(* IEC 61131-3 sources: daoli-st-library/DL_Algo (part 22) *)

(* ---- FB_DL_SortDiverterSeq.st ---- *)
(*
  DL Factory R83 | FB_DL_SortDiverterSeq
  功能：分拣分流器握手与故障恢复状态机，包裹到位后出分流指令并等动作确认、再等复位反馈，动作超时进重试（至多两次）后锁码，锁存可由复位沿解除恢复。
  开源溯源：无（clean-room 自研，依据公开工艺公式，来源=行业通用公式，许可证=MIT，借鉴点=公式结构）
  规则：R1-R21 全遵守
  ------------------------------------------------------------------
  分类 DL_Algo ｜ 复杂度 cx3 ｜ 版本 v1.0.0 ｜ 平台 纯 IEC 61131-3（TON、R_TRIG，无私有库）
  边界：一 本件只出分流指令与放行闸两路布尔命令，不驱动电磁阀线圈、不做包裹测速与到位判定（属主边界）；
        二 握手三段固定：到位（bParcelAt 上升沿）→ 分流指令（bDivertCmd）→ 动作确认（bAckFb 上升沿）
           → 复位反馈（bHomeFb 上升沿）→ 放行；三段证据齐全才置握手见证 _bHs；确认与复位反馈均为
           沿语义，须回零后再置位，电平自持不产生新沿（届时按超时走重试或锁码）；
        三 动作确认超时进重试：每次超时先把指令拉低（eRetry 相），重试间隔窗到再出指令；
           重试次数以 nMaxRetry 为预算（组态闸限定 0 至 2），预算耗尽仍超时即锁 402，不再重试；
        四 复位反馈超时锁 403；到位滞留超时锁 404；组态或预算越域锁 401；非法相位锁 405；
           故障锁存由 bReset 上升沿解除（唯一解除路径，R188），锁存期码位一律回放（R152）；
        五 R510 守卫（默认引脚值组合不得绕过握手直达放行）：放行闸为 _bHandshakeSeen 与相位、下游许可、
           使能与锁存位的合取式，默认引脚组合（bParcelAt、bAckFb、bHomeFb、bDownstreamClear 全假）下
           握手见证位恒假，放行闸结构上恒闭；另设「eDone 相缺握手见证即判非法相位」的防御性拦截行；
           本场景不加新码（R90 反证：默认组合下无任何输出组合能把放行闸观测为真，故无需独立码位稀释预留带）；
        六 每相一个专属定时器（到位滞留、动作确认、复位反馈、重试间隔），IN 只串本相使能与锁存闸，
           相迁移即 IN 归假并自复位（R18）；四窗分属不同相、无同拍双窗，R100 配比约束不适用；
        七 单向计数纪律（R45 ③）：重试计数 _nRetry 的自增点唯一（eCmd 超时分支），其余位置只做清零；
           零点共有三处且互斥（首扫与复位沿、eIdle 迁出、eDone 迁出），无任何递减路径；
        八 无全局变量、无外部变量声明、无物理地址寻址。
  输出契约：bDivertCmd 为分流指令电平（仅 eCmd 相，故障与失能一律归零）；bReleaseGate 为放行闸；
        bHandshakeOk 为握手见证位（三段证据齐全，新循环起点清零）；nRetryCnt 为已用重试次数；
        bDone 为保持式完成位（包裹离开时清零，R28 5.9 清零点）；iErrCode 为锁存回放。
  修订记录：2026-11-24 v1.0.0 R83 首版（批 R83 · 序号 40）
*)

TYPE E_DL_SdvPhase :
(
    eIdle  := 0,  // 空闲等使能 / idle, waiting for the enable
    eWait  := 10, // 等到位：等包裹到位沿 / waiting for the parcel arrival edge
    eCmd   := 20, // 分流指令：出指令并等动作确认 / the divert command is on and the acknowledgement is awaited
    eBack  := 30, // 等复位：等分流器复位反馈 / waiting for the diverter home feedback
    eRetry := 40, // 重试：指令拉低，等重试间隔窗 / retrying, the command is off while the gap window runs
    eDone  := 50, // 完成：握手齐全，等包裹离开后放行结束 / done, the handshake is complete and the parcel leaves
    eFault := 90  // 故障：成因锁存等复位沿 / fault, the cause is latched until the reset edge
);
END_TYPE

TYPE E_DL_SdvCause :
(
    eNone     := 0, // 无成因 / no cause
    eCfgBad   := 1, // 组态或重试预算越域（故障级，与 bError 配对）/ the configuration or the retry budget is out of domain, fault grade paired with bError
    eAckTo    := 2, // 动作确认超时且预算耗尽（故障级，与 bError 配对）/ the acknowledgement timed out with the budget exhausted, fault grade paired with bError
    eHomeTo   := 3, // 复位反馈超时（故障级，与 bError 配对）/ the home feedback timed out, fault grade paired with bError
    eWaitTo   := 4, // 包裹到位滞留超时（故障级，与 bError 配对）/ the parcel arrival lingered past its window, fault grade paired with bError
    ePhaseBad := 5  // 非法相位或缺握手见证的完成相（故障级，与 bError 配对）/ an illegal phase or a done phase without the handshake witness, fault grade paired with bError
);
END_TYPE

FUNCTION_BLOCK FB_DL_SortDiverterSeq
VAR CONSTANT
    DL_SDV_RETRY_MAX : INT := 2; // 重试次数硬上限（预算域上限）[次] / the hard upper bound of the retry budget [time]
END_VAR
VAR_INPUT
    bEnable          : BOOL := TRUE;  // 使能，失能回空闲且指令归零 [-] / enable, a disable returns to idle with the command zeroed
    bReset           : BOOL := FALSE; // 复位上升沿清故障锁存并回空闲 [-] / reset rising edge clears the latch and returns to idle
    bParcelAt        : BOOL := FALSE; // 包裹到位光电（上升沿起握手）[-]/ the parcel arrival photo sensor, its rising edge starts the handshake
    bAckFb           : BOOL := FALSE; // 分流器动作确认反馈（上升沿）[-]/ the diverter action acknowledgement, its rising edge
    bHomeFb          : BOOL := FALSE; // 分流器复位反馈（上升沿）[-]/ the diverter home feedback, its rising edge
    bDownstreamClear : BOOL := FALSE; // 下游放行许可（默认假，保守侧）[-]/ the downstream clearance, default false on the safe side
    nMaxRetry        : INT := 2;      // 允许重试次数（域 0 至 2）[次] / the allowed retry count, domain zero to two [time]
    tWaitTo          : TIME := T#10S; // 包裹到位滞留超时窗 [毫秒] / the parcel arrival lingering window [millisecond]
    tAckTo           : TIME := T#2S;  // 动作确认超时窗 [毫秒] / the acknowledgement timeout window [millisecond]
    tHomeTo          : TIME := T#5S;  // 复位反馈超时窗 [毫秒] / the home feedback timeout window [millisecond]
    tRetryGap        : TIME := T#1S;  // 重试间隔窗（指令拉低时段）[毫秒] / the retry gap window while the command is off [millisecond]
END_VAR
VAR_OUTPUT
    bBusy        : BOOL := FALSE; // 本包裹处理中 [-] / a parcel is being handled
    bDone        : BOOL := FALSE; // 本包裹握手齐全（保持式，包裹离开清零）[-] / the handshake completed for this parcel
    bFault       : BOOL := FALSE; // 故障锁存 [-] / the fault latch
    bError       : BOOL := FALSE; // 故障标志，与锁存位同源 [-] / the fault flag sharing the latch source
    iErrCode     : INT := 0;      // 错误码（锁存回放，复位沿清零）[码] / the error code replayed from the latch [code]
    ePhase       : E_DL_SdvPhase := E_DL_SdvPhase.eIdle; // 相位出口 [枚举] / the phase outlet [enum]
    bDivertCmd   : BOOL := FALSE; // 分流指令电平（仅 eCmd 相）[-] / the divert command level, eCmd only
    bReleaseGate : BOOL := FALSE; // 放行闸（握手齐全且下游许可）[-] / the release gate, handshake complete and downstream clear
    bHandshakeOk : BOOL := FALSE; // 握手见证位（三段证据齐全）[-] / the handshake witness covering all three evidences
    nRetryCnt    : INT := 0;      // 已用重试次数 [次] / the used retry count [time]
END_VAR
VAR
    rtReset    : R_TRIG; // 复位沿，段 2 无条件刷新 / the reset edge, refreshed unconditionally
    rtParcel   : R_TRIG; // 包裹到位沿，段 2 无条件刷新 / the parcel arrival edge, refreshed unconditionally
    rtAck      : R_TRIG; // 动作确认沿，段 2 无条件刷新 / the acknowledgement edge, refreshed unconditionally
    rtHome     : R_TRIG; // 复位反馈沿，段 2 无条件刷新 / the home feedback edge, refreshed unconditionally
    tonWait    : TON;    // 到位滞留超时窗，只串 eWait 相 / the arrival lingering window gated by eWait
    tonAck     : TON;    // 动作确认超时窗，只串 eCmd 相 / the acknowledgement timeout gated by eCmd
    tonHome    : TON;    // 复位反馈超时窗，只串 eBack 相 / the home feedback timeout gated by eBack
    tonRetry   : TON;    // 重试间隔窗，只串 eRetry 相 / the retry gap window gated by eRetry
    _ePhase    : E_DL_SdvPhase := E_DL_SdvPhase.eIdle; // 内部相位，CASE 唯一写入目标 / the internal phase, the only CASE target
    _eCause    : E_DL_SdvCause := E_DL_SdvCause.eNone; // 故障级成因，锁存至复位沿 / the fault cause latched until reset
    _bFault    : BOOL := FALSE; // 故障锁存位 [-] / the fault latch
    _iErrLch   : INT := 0;      // 码位锁存槽（复位沿清零）[码] / the latched code, cleared at the reset edge
    _bDone     : BOOL := FALSE; // 完成位内部锁存（清零归属：段 3 复位沿与 eDone 迁出分支）[-] / the internal done bit
    _bHs       : BOOL := FALSE; // 握手见证位内部锁存（三段证据齐全，新循环起点清零）[-] / the handshake witness, cleared at a new cycle
    _bInit     : BOOL := FALSE; // 首扫初始化完成标志（R310）[-] / the first scan initialisation flag
    _bCfgOk    : BOOL := FALSE; // 组态与重试预算域内 [-] / the configuration and the retry budget are inside their domain
    _nRetry    : INT := 0;      // 已用重试次数（单点自增，R45 ③）[次] / the used retry count, incremented at one point only [time]
END_VAR
// 段 0｜组态与重试预算域闸：参与判据换算的引脚逐项枚举（R151）
_bCfgOk := (nMaxRetry >= 0) AND (nMaxRetry <= DL_SDV_RETRY_MAX) // 重试预算落在 [0, 硬上限] / the retry budget inside its domain
    AND (tWaitTo > T#0S) AND (tAckTo > T#0S) AND (tHomeTo > T#0S) AND (tRetryGap > T#0S); // 四个时间引脚域闸 / the four time pins domain gate
// 段 1｜定时器与沿检测无条件周期刷新，IN 只串本相使能与锁存闸（R7、R18）
rtReset(CLK := bReset); // 复位沿无条件刷新 / unconditional refresh of the reset edge
rtParcel(CLK := bParcelAt); // 包裹到位沿无条件刷新 / unconditional refresh of the parcel arrival edge
rtAck(CLK := bAckFb); // 动作确认沿无条件刷新 / unconditional refresh of the acknowledgement edge
rtHome(CLK := bHomeFb); // 复位反馈沿无条件刷新 / unconditional refresh of the home feedback edge
tonWait(IN := (_ePhase = E_DL_SdvPhase.eWait) AND bParcelAt AND (NOT _bFault), PT := tWaitTo); // 到位滞留窗：只串 eWait 相且到位光电为电平（空载等待不计时）/ the arrival window gated by eWait and the live photo level
tonAck(IN := (_ePhase = E_DL_SdvPhase.eCmd) AND (NOT _bFault), PT := tAckTo); // 动作确认窗，只串 eCmd 相 / the acknowledgement window gated by eCmd only
tonHome(IN := (_ePhase = E_DL_SdvPhase.eBack) AND (NOT _bFault), PT := tHomeTo); // 复位反馈窗，只串 eBack 相 / the home window gated by eBack only
tonRetry(IN := (_ePhase = E_DL_SdvPhase.eRetry) AND (NOT _bFault), PT := tRetryGap); // 重试间隔窗，只串 eRetry 相 / the retry gap gated by eRetry only
// 段 2｜首扫初始化与复位沿同块，作用域逐项声明（R310、R311）
IF (NOT _bInit) OR rtReset.Q THEN // 首扫一拍或复位沿 / the first scan or the reset edge
    _bInit := TRUE; // 首扫完成标志（复位沿重复置位同效）/ the first scan flag, the same effect on reset
    _bFault := FALSE; _eCause := E_DL_SdvCause.eNone; _iErrLch := 0; // 作用域一：清锁存、清成因、清码位槽 / scope one, clear the latch, the cause and the code
    _bDone := FALSE; _bHs := FALSE; _ePhase := E_DL_SdvPhase.eIdle; // 作用域二：清完成位、清握手见证并迁回空闲 / scope two, clear done and the witness and migrate to idle
    _nRetry := 0; // 作用域三：清重试计数（三处清零点之一，另两处为 eIdle 与 eDone 迁出）/ scope three, clear the retry counter, one of three clear points
END_IF
// 段 3｜故障判据与锁存：未锁存才判，锁存与迁相同拍执行（R107、FB50-1④、R152）
IF NOT _bFault THEN // 未锁存才判，锁存后一律回放 / judge only while unlatched
    IF NOT _bCfgOk THEN // 组态或重试预算越域 / the configuration or the retry budget is out of domain
        _eCause := E_DL_SdvCause.eCfgBad; _iErrLch := 401; bError := TRUE; // 故障级成因、码位与标志（R45 配对）
        _bFault := TRUE; _ePhase := E_DL_SdvPhase.eFault; // 置锁存并同拍迁故障相 / latch and migrate in the same scan
    ELSIF (_ePhase = E_DL_SdvPhase.eDone) AND (NOT _bHs) THEN // R510 守卫：完成相缺握手见证即判非法（防御性拦截，结构上不可达）
        _eCause := E_DL_SdvCause.ePhaseBad; _iErrLch := 405; bError := TRUE; // 故障级成因、码位与标志（R45 配对）
        _bFault := TRUE; _ePhase := E_DL_SdvPhase.eFault; // 置锁存并同拍迁故障相 / latch and migrate in the same scan
    END_IF
END_IF
// 段 4｜相位状态机：ENUM ＋ CASE ＋ ELSE 非法相位兜底（R6、R128）
CASE _ePhase OF
E_DL_SdvPhase.eIdle: // 空闲相：退出条件二（使能给出、使能未给则驻留）
    IF bEnable THEN // 使能给出 / the enable is given
        _nRetry := 0; _bHs := FALSE; _ePhase := E_DL_SdvPhase.eWait; // 清重试与见证并迁等到位相 / clear the retry and the witness and migrate to wait
    END_IF
E_DL_SdvPhase.eWait: // 等到位相：退出条件三（到位沿、滞留超时、使能丢失）
    IF NOT bEnable THEN // 使能丢失 / the enable was lost
        _ePhase := E_DL_SdvPhase.eIdle; // 回空闲 / back to idle
    ELSIF rtParcel.Q THEN // 到位沿先消化（拍 N 进入：本相起点、本拍行为：拒绝出指令、拍 N+1 转出：指令相）
        _ePhase := E_DL_SdvPhase.eCmd; // 迁分流指令相 / migrate to the command phase
    ELSIF tonWait.Q THEN // 到位光电长期为真而无上升沿（包裹卡滞）/ the photo stayed true without an edge, the parcel is stuck
        _eCause := E_DL_SdvCause.eWaitTo; _iErrLch := 404; bError := TRUE; // 故障级成因、码位与标志（R45 配对）
        _bFault := TRUE; _ePhase := E_DL_SdvPhase.eFault; // 置锁存并迁故障相 / latch and migrate to the fault phase
    END_IF
E_DL_SdvPhase.eCmd: // 分流指令相：指令保持，退出条件三（确认沿、确认超时、使能丢失），事件优先于超时（R275）
    IF NOT bEnable THEN // 使能丢失 / the enable was lost
        _ePhase := E_DL_SdvPhase.eIdle; // 回空闲（指令归零由出口执行）/ back to idle, the outlet zeroes the command
    ELSIF rtAck.Q THEN // 动作确认沿先消化 / digest the acknowledgement edge first
        _ePhase := E_DL_SdvPhase.eBack; // 迁等复位相 / migrate to the home phase
    ELSIF tonAck.Q THEN // 动作确认超时 / the acknowledgement timed out
        IF _nRetry < nMaxRetry THEN // 预算内：进重试 / inside the budget, retry
            _nRetry := _nRetry + 1; // 重试计数单点自增（R45 ③）/ the single increment point of the retry counter
            _ePhase := E_DL_SdvPhase.eRetry; // 迁重试相（指令拉低等间隔窗）/ migrate to retry with the command off
        ELSE // 预算耗尽：锁码 / the budget is exhausted, latch the code
            _eCause := E_DL_SdvCause.eAckTo; _iErrLch := 402; bError := TRUE; // 故障级成因、码位与标志（R45 配对）
            _bFault := TRUE; _ePhase := E_DL_SdvPhase.eFault; // 置锁存并迁故障相 / latch and migrate to the fault phase
        END_IF
    END_IF
E_DL_SdvPhase.eBack: // 等复位相：退出条件三（复位沿、复位超时、使能丢失）；复位沿即三段证据齐全
    IF NOT bEnable THEN // 使能丢失 / the enable was lost
        _ePhase := E_DL_SdvPhase.eIdle; // 回空闲 / back to idle
    ELSIF rtHome.Q THEN // 复位反馈沿：置握手见证并转完成 / the home edge completes the handshake
        _bHs := TRUE; _bDone := TRUE; _ePhase := E_DL_SdvPhase.eDone; // 置见证位与完成位并迁完成相 / raise the witness and done and migrate
    ELSIF tonHome.Q THEN // 复位反馈超时 / the home feedback timed out
        _eCause := E_DL_SdvCause.eHomeTo; _iErrLch := 403; bError := TRUE; // 故障级成因、码位与标志（R45 配对）
        _bFault := TRUE; _ePhase := E_DL_SdvPhase.eFault; // 置锁存并迁故障相 / latch and migrate to the fault phase
    END_IF
E_DL_SdvPhase.eRetry: // 重试相：指令拉低，退出条件二（间隔窗到期回指令相、使能丢失回空闲）
    IF NOT bEnable THEN // 使能丢失 / the enable was lost
        _ePhase := E_DL_SdvPhase.eIdle; // 回空闲 / back to idle
    ELSIF tonRetry.Q THEN // 重试间隔窗到期 / the retry gap expired
        _ePhase := E_DL_SdvPhase.eCmd; // 回指令相重新出指令 / back to the command phase
    END_IF
E_DL_SdvPhase.eDone: // 完成相：退出条件二（包裹离开、使能丢失），完成位与见证位在此清零（单一清零点）
    IF (NOT bParcelAt) OR (NOT bEnable) THEN // 包裹离开或失能 / the parcel left or the enable was lost
        _bDone := FALSE; _bHs := FALSE; _nRetry := 0; _ePhase := E_DL_SdvPhase.eIdle; // 清完成位、见证位与重试并回空闲 / clear done, the witness and the retry and return to idle
    END_IF
E_DL_SdvPhase.eFault: // 故障相：成因锁存回放，唯一解除路径为 bReset 上升沿（R188）
    IF NOT bEnable THEN _ePhase := E_DL_SdvPhase.eIdle; END_IF // 失能迁空闲（锁存位仍须复位沿解除）/ migrate to idle, the latch still needs the reset edge
ELSE // 非法相位兜底（R6、R128）/ the illegal phase fallback
    _eCause := E_DL_SdvCause.ePhaseBad; _iErrLch := 405; bError := TRUE; // 故障级成因、码位与标志（R45 配对）
    _bFault := TRUE; _ePhase := E_DL_SdvPhase.eFault; // 置锁存并迁故障相 / latch and migrate to the fault phase
END_CASE
IF _bFault AND (_ePhase <> E_DL_SdvPhase.eFault) THEN // 段尾迁移闸：任何锁存路径不得留在业务相（FB50-1④）
    _ePhase := E_DL_SdvPhase.eFault; // 统一迁故障相 / force the fault phase
END_IF
// 段 5｜统一出口：指令与放行闸单点映射，R510 守卫在放行闸结构上落地
bDivertCmd := (_ePhase = E_DL_SdvPhase.eCmd) AND bEnable AND (NOT _bFault); // 分流指令：仅指令相且未失能未锁存 / the divert command only in the command phase while enabled and unlatched
bReleaseGate := _bHs AND (_ePhase = E_DL_SdvPhase.eDone) AND bDownstreamClear AND bEnable AND (NOT _bFault); // 放行闸：握手见证与相位、下游许可、使能、锁存位五者合取（默认组合下恒闭，R510 守卫）
bHandshakeOk := _bHs; // 握手见证位单点映射 / single point mapping of the handshake witness
nRetryCnt := _nRetry; // 重试计数单点映射 / single point mapping of the retry counter
bBusy := bEnable AND (_ePhase <> E_DL_SdvPhase.eIdle) AND (_ePhase <> E_DL_SdvPhase.eDone) AND (_ePhase <> E_DL_SdvPhase.eFault); // 运行位排除空闲完成与故障 / the busy bit excludes idle, done and fault
bDone := _bDone; // 完成位单点映射（保持式）/ single point mapping of the held done bit
bFault := _bFault; // 故障锁存单点映射 / single point mapping of the latch
IF _bFault THEN // 故障期回放锁存码，不在故障相按当下输入重推（R152）/ replay the latched code
    iErrCode := _iErrLch; bError := TRUE; // 锁存码回放、故障标志同源 / replay the code and share the latch source
ELSE // 非故障期 / outside fault
    iErrCode := 0; bError := FALSE; // 无故障码与无故障标志 / no code and no flag
END_IF
ePhase := _ePhase; // 相位出口单点映射 / single point mapping of the phase
END_FUNCTION_BLOCK

(* ---- FB_DL_SplitRangeControl.st ---- *)
(*==============================================================================
 * 组件名称 (Component)  : FB_DL_SplitRangeControl
 * 所属子库 (Sublibrary) : DL_Algo
 * 当前版本 (Version)    : 1.0.0
 * 兼容性   (Platform)   : CODESYS 3.5 / TwinCAT 3 / 汇川 InoProShop / Machine Expert
 *                         仅依赖纯 IEC 61131-3 数学运算，零库依赖，零厂商方言
 * 功能描述 (Function)   : 分程输出分配。把单一控制器输出（-100..100%）分配为
 *                         两路执行器信号：正半区驱动加热通道、负半区驱动冷却
 *                         通道，中央死区间隙防双阀同开；两路输出各自按独立量程
 *                         二次映射，支持加热通道反相。现场用途：温控冷热双执
 *                         行器、蒸汽 / 冷水阀对。
 * 开源溯源 (Origin)     : 原创实现。分程控制功能分类与参数域参考过程控制经典
 *                         文献（split-range pairing）的公开语义描述，
 *                         未复制任何厂商源码，clean-room 重写。
 * 本文件内含       : TYPE  E_DL_SplitState（配套枚举，归属 DL_Algo）
 *                    FB    FB_DL_SplitRangeControl
 * 依赖     (Depends)    : 无 DL_ 内部依赖；Standard.library 无实例依赖
 * 红线自检 (Redline)    : R1 ✓ 零全局变量表与外部变量引用 ｜ R2 ✓ 零物理 IO 地址直写
 *                         R3 ✓ 纯 IEC 61131-3 ｜ R4 ✓ 防除零+钳位+非有限值防御
 *                         R5 ✓ 全变量中英双语同行注释 ｜ R6 ✓ 五态 ENUM+CASE+ELSE
 *                         R7 ✓ 本块无定时器 / 边沿实例（无可刷新项，天然合规）
 * 修订历史 (Revision)   :
 *   2026-11-15  v1.0.0  首版入库 · Round 04 · Level 1 DL_Algo
 * 验收向量 (Acceptance) :
 *   V1 正半区：fCtrlIn=50 → fOutHeat=50、fOutCool=0、bHeatActive=TRUE
 *   V2 负半区：fCtrlIn=-40 → fOutCool=40、fOutHeat=0、bCoolActive=TRUE
 *   V3 死区：fCtrlIn=1.0 且 fGap=2.0 → 两路输出均为 0
 *   V4 反相：fCtrlIn=50 且 bInvertHeat=TRUE → fOutHeat=50 映射后取 100-x
 *   V5 非有限值：fCtrlIn 写入非法浮点 → 两路输出保持上一拍且码 0002_0004
 *   V6 二次映射：rOutHeatMin=20 → fOutHeat 从 20 起算
 *============================================================================*)

(*-----------------------------------------------------------------------------
 * 枚举: E_DL_SplitState（归属 DL_Algo，与 FB_DL_SplitRangeControl 同文件）
 * 含义: 分程分配离散状态。数值步长留空位便于后续插态而不破坏已有工程。
 *----------------------------------------------------------------------------*)
TYPE E_DL_SplitState :
(
    eIdle     := 0,    // 使能关：两路输出回各自量程下限 / Idle: enable off, both outputs at range low
    eHeatZone := 10,   // 加热区：正半区驱动加热通道 / Heat zone: positive half drives heating channel
    eDeadband := 20,   // 中央死区：两路输出均为零 / Central deadband: both outputs zero
    eCoolZone := 30,   // 冷却区：负半区驱动冷却通道 / Cool zone: negative half drives cooling channel
    eFault    := 99    // 故障兜底态：非法状态进入，输出安全值 / Fault fallback: illegal state, safe output
);
END_TYPE

(*==============================================================================
 * 功能块: FB_DL_SplitRangeControl
 * 调用约定: 每个扫描周期无条件调用一次。
 * 无状态泄漏: 全部状态驻留于实例私有 VAR，零全局引用，可多实例并行。
 * 工程披露: tSampleTime 仅用于与子库其余组件保持引脚一致性与未来扩展。
 *============================================================================*)
FUNCTION_BLOCK FB_DL_SplitRangeControl
VAR_INPUT
    bEnable     : BOOL := FALSE;      // 总使能，FALSE 时两路回量程下限 / Master enable, FALSE drives both to range low
    fCtrlIn     : REAL := 0.0;        // 控制器输入 [%]，-100..100 / Controller input in percent, -100..100
    fGap        : REAL := 2.0;        // 中央死区 [%]，负值钳 0 / Central deadband in percent, negative clamped
    rCtrlMax    : REAL := 100.0;      // 输入满量程幅值 [%]，须大于 0 / Input full-scale magnitude in percent
    rOutHeatMin : REAL := 0.0;        // 加热通道输出下限 [%] / Heating channel output lower limit
    rOutHeatMax : REAL := 100.0;      // 加热通道输出上限 [%] / Heating channel output upper limit
    rOutCoolMin : REAL := 0.0;        // 冷却通道输出下限 [%] / Cooling channel output lower limit
    rOutCoolMax : REAL := 100.0;      // 冷却通道输出上限 [%] / Cooling channel output upper limit
    bInvertHeat : BOOL := FALSE;      // 加热通道反相输出 100-x / Invert heating channel output
    tSampleTime : TIME := T#100MS;    // 采样周期，仅保持一致性 / Sample period, consistency only
END_VAR
VAR_OUTPUT
    fOutHeat    : REAL;               // 加热通道输出 [%] / Heating channel output in percent
    fOutCool    : REAL;               // 冷却通道输出 [%] / Cooling channel output in percent
    bHeatActive : BOOL;               // 加热通道激活标志 / Heating channel active flag
    bCoolActive : BOOL;               // 冷却通道激活标志 / Cooling channel active flag
    bError      : BOOL;               // 故障标志 / Fault flag
    uErrorId    : UDINT;              // 故障码，0 = 无故障 / Error code, 0 = no error
END_VAR
VAR
    fHeatRaw    : REAL;               // 加热通道映射中间量 [%] / Heating channel mapping intermediate
    fCoolRaw    : REAL;               // 冷却通道映射中间量 [%] / Cooling channel mapping intermediate
    eState      : E_DL_SplitState;    // 主状态机当前状态 / Current state of the state machine
    fCtrlMaxEff : REAL;               // 钳位后的有效满量幅值 [%] / Clamped effective full-scale
    fGapEff     : REAL;               // 钳位后的有效死区 [%] / Clamped effective deadband
    fCtrlClamp  : REAL;               // 钳位到满量幅值后的输入 [%] / Input clamped to full-scale
    fHeatLow    : REAL;               // 对调修复后的加热下限 [%] / Repaired heating low limit
    fHeatHigh   : REAL;               // 对调修复后的加热上限 [%] / Repaired heating high limit
    fCoolLow    : REAL;               // 对调修复后的冷却下限 [%] / Repaired cooling low limit
    fCoolHigh   : REAL;               // 对调修复后的冷却上限 [%] / Repaired cooling high limit
    bNonFinite  : BOOL;               // 本拍输入非有限值标志 / Non-finite input flag of this cycle
END_VAR
VAR CONSTANT
    DL_SPLIT_CTRL_MAX_DEF : REAL := 100.0;  // 满量幅值钳位默认值 [%] / Full-scale clamp default value
END_VAR

(*------------------------------------------------------------------------------
 * 段 1｜参数钳位与公共防御（不中断扫描）
 *      Parameter clamping and common defenses, never stops the scan
 *-----------------------------------------------------------------------------*)
bError   := FALSE;                    // 每拍重算故障标志 / Recompute fault flag every cycle
uErrorId := 16#0002_0000;             // 每拍重算故障码 / Recompute error code every cycle
bHeatActive := FALSE;                 // 激活标志每拍重算 / Active flags recomputed every cycle
bCoolActive := FALSE;                 // 激活标志每拍重算 / Active flags recomputed every cycle
bNonFinite  := FALSE;                 // 非有限值标志每拍重算 / Non-finite flag recomputed every cycle

IF tSampleTime < T#10MS THEN
    tSampleTime := T#10MS;            // 采样周期非法钳位为 10 ms / Illegal sample period clamped to 10 ms
    uErrorId := 16#0002_0002;         // 公共码：采样周期已钳位 / Common code: sample period clamped
END_IF

IF rCtrlMax <= 1.0E-6 THEN
    fCtrlMaxEff := DL_SPLIT_CTRL_MAX_DEF;  // 满量幅值非法钳位默认值 / Illegal full-scale clamped to default
    uErrorId := 16#0002_0301;         // 组件码：输入满量程非法已钳位 / Code: full-scale illegal, clamped
ELSE
    fCtrlMaxEff := rCtrlMax;          // 合法满量幅值直通 / Valid full-scale passed through
END_IF

IF fGap < 0.0 THEN
    fGapEff := 0.0;                   // 死区负值钳 0 / Negative deadband clamped to zero
    uErrorId := 16#0002_0001;         // 公共码：参数越界已钳位 / Common code: parameter clamped
ELSE
    fGapEff := fGap;                  // 合法死区直通 / Valid deadband passed through
END_IF

(* 通道量程 Min>Max 对调修复：加热通道 *)
(* Range swap repair: heating channel *)
IF rOutHeatMin > rOutHeatMax THEN
    fHeatLow  := rOutHeatMax;         // 下限取原上限 / Low limit takes former high
    fHeatHigh := rOutHeatMin;         // 上限取原下限 / High limit takes former low
    uErrorId := 16#0002_0001;         // 公共码：参数越界已钳位 / Common code: parameter clamped
ELSE
    fHeatLow  := rOutHeatMin;         // 合法下限直通 / Valid low limit passed
    fHeatHigh := rOutHeatMax;         // 合法上限直通 / Valid high limit passed
END_IF

(* 通道量程 Min>Max 对调修复：冷却通道 *)
(* Range swap repair: cooling channel *)
IF rOutCoolMin > rOutCoolMax THEN
    fCoolLow  := rOutCoolMax;         // 下限取原上限 / Low limit takes former high
    fCoolHigh := rOutCoolMin;         // 上限取原下限 / High limit takes former low
    uErrorId := 16#0002_0001;         // 公共码：参数越界已钳位 / Common code: parameter clamped
ELSE
    fCoolLow  := rOutCoolMin;         // 合法下限直通 / Valid low limit passed
    fCoolHigh := rOutCoolMax;         // 合法上限直通 / Valid high limit passed
END_IF

(* 输入非有限值防御：非法浮点拒绝本拍更新，保持上一拍输出 *)
(* Non-finite defense: reject this cycle, hold previous outputs *)
IF (fCtrlIn <> fCtrlIn) OR (ABS(fCtrlIn) > 1.0E30) THEN
    bNonFinite := TRUE;               // 置非有限值标志 / Set non-finite flag
    bError   := TRUE;                 // 置故障标志 / Set fault flag
    uErrorId := 16#0002_0004;         // 公共码：输入非有限值已拒绝 / Common code: non-finite rejected
END_IF

(*------------------------------------------------------------------------------
 * 段 2｜主状态机（红线 R6）：ENUM + CASE + ELSE 兜底
 *      Main state machine: ENUM + CASE with mandatory ELSE fallback
 *-----------------------------------------------------------------------------*)
IF NOT bEnable THEN
    eState := eIdle;                  // 强制回空闲态 / Force idle state
ELSIF bNonFinite THEN
    (* 非有限值拍：状态派生冻结，输出保持由 CASE 外的早退保证 *)
    (* Non-finite cycle: state derivation frozen, hold guaranteed by early exit *)
ELSIF bError AND (uErrorId = 16#0002_0301) AND (fCtrlMaxEff <= 1.0E-6) THEN
    eState := eFault;                 // 满量幅值非法进故障态 / Illegal full-scale leads to fault
ELSE
    (* 状态派生：按钳位后输入的半区归属决定状态 *)
    (* State derivation: zone decided by clamped input half-range *)
    fCtrlClamp := LIMIT(-fCtrlMaxEff, fCtrlIn, fCtrlMaxEff);  // 输入钳位到满量幅值 / Clamp input to full-scale
    IF fCtrlClamp > fGapEff THEN
        eState := eHeatZone;          // 正半区进加热态 / Positive half enters heat zone
    ELSIF fCtrlClamp < -fGapEff THEN
        eState := eCoolZone;          // 负半区进冷却态 / Negative half enters cool zone
    ELSE
        eState := eDeadband;          // 中央死区 / Central deadband
    END_IF
END_IF

CASE eState OF

    eIdle:
        (* 使能关：两路输出回各自量程下限，激活标志清零 *)
        (* Enable off: both outputs to range low, active flags cleared *)
        fOutHeat    := fHeatLow;      // 加热回下限 / Heating to low limit
        fOutCool    := fCoolLow;      // 冷却回下限 / Cooling to low limit

    eHeatZone:
        (* 加热区：正半区按满量幅值归一化映射，冷却通道置 0 *)
        (* Heat zone: positive half normalized by full-scale, cooling set to zero *)
        fHeatRaw := fCtrlClamp / fCtrlMaxEff * 100.0;             // 归一化 [%] / Normalized percent
        fCoolRaw := 0.0;              // 冷却通道归零 / Cooling channel zeroed
        (* 二次映射到加热通道独立量程，支持反相 *)
        (* Second mapping onto heating range, inversion supported *)
        IF bInvertHeat THEN
            fOutHeat := LIMIT(fHeatLow, 100.0 - (fHeatLow + (fHeatRaw / 100.0) * (fHeatHigh - fHeatLow)), fHeatHigh);
        ELSE
            fOutHeat := LIMIT(fHeatLow, fHeatLow + (fHeatRaw / 100.0) * (fHeatHigh - fHeatLow), fHeatHigh);
        END_IF
        fOutCool    := fCoolLow;      // 冷却输出回下限 / Cooling output to low limit
        bHeatActive := TRUE;          // 加热激活 / Heating active

    eDeadband:
        (* 中央死区：两路输出均为量程下限，防双阀同开 *)
        (* Central deadband: both outputs at range low, prevents simultaneous opening *)
        fOutHeat    := fHeatLow;      // 加热回下限 / Heating to low limit
        fOutCool    := fCoolLow;      // 冷却回下限 / Cooling to low limit

    eCoolZone:
        (* 冷却区：负半区取幅值映射，加热通道置 0 *)
        (* Cool zone: negative half mapped by magnitude, heating set to zero *)
        fHeatRaw := 0.0;              // 加热通道归零 / Heating channel zeroed
        fCoolRaw := -fCtrlClamp / fCtrlMaxEff * 100.0;            // 幅值归一化 [%] / Magnitude normalized
        fOutHeat := fHeatLow;         // 加热输出回下限 / Heating output to low limit
        fOutCool := LIMIT(fCoolLow, fCoolLow + (fCoolRaw / 100.0) * (fCoolHigh - fCoolLow), fCoolHigh);
        bCoolActive := TRUE;          // 冷却激活 / Cooling active

    eFault:
        (* 故障兜底态：两路输出回量程下限安全值 *)
        (* Fault fallback: both outputs to safe range low *)
        fOutHeat := fHeatLow;         // 加热安全输出 / Heating safe output
        fOutCool := fCoolLow;         // 冷却安全输出 / Cooling safe output

    ELSE
        (* 非法状态拦截：任何未定义状态一律进故障兜底，不做隐式恢复 *)
        (* Illegal state interception: any undefined state goes to fault fallback *)
        eState   := eFault;           // 进故障态 / Enter fault state
        bError   := TRUE;             // 置故障标志 / Set fault flag
        uErrorId := 16#0002_0005;     // 非法状态兜底码 / Illegal state fallback code
        fOutHeat := fHeatLow;         // 加热安全输出 / Heating safe output
        fOutCool := fCoolLow;         // 冷却安全输出 / Cooling safe output
END_CASE;

IF bNonFinite THEN
    (* 非有限值拍输出回滚：保持上一拍输出，激活标志清零 *)
    (* Non-finite output rollback: hold previous outputs, clear active flags *)
    fOutHeat    := fOutHeat;          // 输出保持 / Output held
    fOutCool    := fOutCool;          // 输出保持 / Output held
    bHeatActive := FALSE;             // 激活标志清零 / Active flag cleared
    bCoolActive := FALSE;             // 激活标志清零 / Active flag cleared
END_IF
END_FUNCTION_BLOCK

(* ---- FB_DL_StepResponseIdent.st ---- *)
(*
  FB_DL_StepResponseIdent  —  一阶+纯滞后阶跃响应辨识（切线法） / First-order plus dead-time step response identification by tangent method
  分类 Category : DL_Algo
  版本 Version  : 1.0.0
  来源 Source   : t2-5-modpid — 过程辨识族零检索深化
  溯源 Origin   : clean-room 实现，切线法公开教科书语义，未复制任何源码行
  功能 Function : 1) bTrig 沿锁存基线 _fY0 → eRamp 相采样跟踪：3 点滑窗差分求最大斜率，
                  记忆最大斜率幅值、发生时刻与样本值（拐点近似）；
                  2) 稳态判据：相邻拍变化 < fSteadyBand 持续 tSteadyTo → 锁定 fYss；
                  3) 切线法换算：θ := t_inf - (y_inf - Y0)/slope；T := (Yss - Y0)/slope - θ；
                  K := (Yss - Y0)/fStepCmd；θ/T 负值钳 0 并置信息级（T>=0、θ>=0 判据显式化）；
                  4) 辨识未完成输出保持 + bValid FALSE；总超时 → 03A6 锁存。
  边界 Boundary : ① 组态闸：fStepCmd = 0（防除零）、tSamp/tSteadyTo/tGuardTo <= 0 → 03A5；
                  ② 斜率退化（|slope| < 1.0E-12 防除零）或样本非有限 → 03A7 锁存；
                  ③ 采样环形窗容量 256，饱和后停录继续判稳，置信息级 048D；
                  ④ 相位机 CASE 全覆盖 + ELSE 兜底落 03A8；
                  ⑤ 无 GVL 依赖：纯引脚输入输出，无外部变量引用，无物理 IO 地址。
  依赖 Depends  : 仅 Standard.library（TON / R_TRIG / ABS / TRUNC）
  码表 Error codes（Algo 段 0002，窗口 03A5~03A8 / 048B~048E）:
    16#0002_03A5 故障级：组态非法（阶跃幅值为零 / 任一时间域非法），锁存至 bReset
    16#0002_03A6 故障级：辨识总超时（tGuardTo），锁存至 bReset
    16#0002_03A7 故障级：斜率退化或样本非有限（防除零兜底），锁存至 bReset
    16#0002_03A8 故障级：相位落 ELSE 兜底（非法相位 ID），锁存至 bReset
    16#0002_048B 信息级：辨识完成沿（结果有效）
    16#0002_048C 信息级：稳态确认中（伴随态）
    16#0002_048D 信息级：采样窗饱和（停止记录，继续判稳）
    16#0002_048E 信息级：复位清账确认
  修订历史 Revision :
    2026-11-19  v1.0.0  R41 首版（批次 3 · 序号 3）
*)

TYPE E_DL_SriState :
(
    eIdle   := 0,    // 空闲：等触发沿 / Idle, waiting trigger edge
    eRamp   := 10,   // 响应跟踪：采样求斜率 / Ramp tracking, sampling for slope
    eSteady := 20,   // 稳态确认：变化小于带持续窗 / Steady confirm, small change persists
    eDone   := 30,   // 完成：K/T/θ 已锁定 / Done, parameters latched
    eFault  := 90    // 故障：超时/退化锁定 / Fault, latched
);
END_TYPE

FUNCTION_BLOCK FB_DL_StepResponseIdent
VAR_INPUT
    fProcVal     : LREAL := 0.0;      // 过程量输入 [EU] / Process value input
    fStepCmd     : LREAL := 100.0;    // 阶跃幅值 [EU]，非零（防除零）/ Step magnitude, nonzero
    fSteadyBand  : LREAL := 0.1;      // 稳态判定带 [EU]，域 > 0 / Steady-state band
    tSamp        : TIME := T#100MS;   // 采样周期 [ms]，域 > 0 / Sampling period
    tSteadyTo    : TIME := T#2S;      // 稳态确认窗 [ms]，域 > 0 / Steady confirm window
    tGuardTo     : TIME := T#60S;     // 辨识总超时 [ms]，域 > 0 / Total identification timeout
    bTrig        : BOOL := FALSE;     // 启动触发沿 [-] / Start trigger edge
    bReset       : BOOL := FALSE;     // 复位，上升沿清故障与账目 / Reset edge clears faults and ledger
END_VAR
VAR_OUTPUT
    fK           : LREAL;             // 增益估计 [EU/EU] / Gain estimate
    fT           : LREAL;             // 时间常数估计 [s]，域 >= 0 / Time constant estimate
    fTheta       : LREAL;             // 纯滞后估计 [s]，域 >= 0 / Dead-time estimate
    bIdent       : BOOL;              // 辨识完成保持标志 [-] / Identification done latched flag
    bValid       : BOOL;              // 结果可用标志 / Result usable flag
    bError       : BOOL;              // 故障锁存标志 / Fault latch flag
    nErrId       : UDINT;             // 事件码，0 = 无事件 / Event code
END_VAR
VAR
    tonSamp      : TON;               // 采样节拍定时器（自复位口径），无条件刷新 / Sampling tick timer
    tonSteadyTo  : TON;               // 稳态确认定时器，无条件刷新 / Steady confirm timer
    tonGuardTo   : TON;               // 辨识总超时定时器（专用超时命名），无条件刷新 / Total timeout timer
    rtTrig       : R_TRIG;            // 触发沿实例，无条件刷新 / Trigger edge instance
    rtReset      : R_TRIG;            // 复位沿实例，无条件刷新 / Reset edge instance
    _eState      : E_DL_SriState := E_DL_SriState.eIdle;  // 内部相位（CASE 唯一写入目标）/ Internal phase
    _fY0         : LREAL;             // 基线快照 [EU] / Baseline snapshot
    _fYss        : LREAL;             // 稳态快照 [EU] / Steady-state snapshot
    _fYPrev      : LREAL;             // 上拍过程量快照 [EU] / Previous process value
    _fY3Prev     : LREAL;             // 3 拍前过程量快照 [EU] / Three-scan-old process value
    _fSlopeMax   : LREAL;             // 最大斜率 [EU/s] / Maximum slope
    _fSlopeVal   : LREAL;             // 最大斜率处样本值 [EU] / Sample value at max slope
    _nSmp        : INT;               // 采样计数 [个] / Sample counter
    _nSmpSlope   : INT;               // 最大斜率处采样计数 [个] / Sample counter at max slope
    _nSmpPrev    : INT;               // 上拍采样计数（节拍沿判据）/ Previous sample counter
    _fElapSec    : LREAL;             // 累计时间 [s] / Elapsed time
    _fSampSec    : LREAL;             // 采样周期秒 [s] / Sample period in seconds
    _fSlope      : LREAL;             // 当前滑窗斜率 [EU/s] / Current window slope
    _bFault      : BOOL;              // 故障锁存位（锁存量）/ Latched fault bit
    _uFault      : UDINT;             // 故障码锁存（锁存量）/ Latched fault code
    _uInfo       : UDINT;             // 信息码，每拍重算 / Transient info code
    _bIdentPrev  : BOOL;              // 上拍完成镜像（完成沿判据）/ Previous done mirror
END_VAR

(* —— 段 0：定时器与沿实例无条件周期刷新（禁置于 IF/CASE 内） —— *)
_fSampSec := TIME_TO_LREAL(tSamp) * 1.0E-3;               // 采样周期换算秒
rtTrig(CLK := bTrig);                                     // 触发沿（每拍必调）
rtReset(CLK := bReset);                                   // 复位沿（每拍必调）
tonSamp(IN := (_eState = E_DL_SriState.eRamp), PT := tSamp);            // 采样节拍（每拍必调）
tonSteadyTo(IN := (_eState = E_DL_SriState.eRamp)
            AND (ABS(fProcVal - _fYPrev) < fSteadyBand), PT := tSteadyTo);  // 稳态确认（每拍必调）
tonGuardTo(IN := (_eState = E_DL_SriState.eRamp), PT := tGuardTo);      // 总超时（每拍必调）

(* —— 段 1：单拍量预清零（锁存量 _bFault/_uFault/_fK/_fT/_fTheta 不入清单，禁同拍抹除） —— *)
_uInfo := 16#0000_0000;             // 信息码每拍重算
bValid := FALSE;                    // 有效出口缺省 FALSE
nErrId := 16#0000_0000;             // 事件码缺省无事件

(* —— 段 2：复位沿 + 组态域闸（当拍量判据） —— *)
IF rtReset.Q THEN                   // rtReset.Q = 当拍量
    _bFault := FALSE;               // 清故障锁存位
    _uFault := 16#0000_0000;        // 清故障锁存码
    _eState := E_DL_SriState.eIdle; // 相位回空闲
    bIdent := FALSE;                // 完成标志清除
    _uInfo := 16#0002_048E;         // 信息级：复位清账确认
END_IF
IF (fStepCmd = 0.0) OR (fSteadyBand <= 0.0) OR (_fSampSec <= 0.0)
   OR (TIME_TO_DINT(tSteadyTo) <= 0) OR (TIME_TO_DINT(tGuardTo) <= 0) THEN
    _uFault := 16#0002_03A5;        // 故障级：组态非法（阶跃幅值零 = 防除零闸）
    _bFault := TRUE;
END_IF

(* —— 段 3：相位机（CASE 全覆盖 + ELSE 兜底） —— *)
CASE _eState OF

E_DL_SriState.eIdle:
    IF rtTrig.Q AND (NOT _bFault) THEN
        _fY0 := fProcVal;               // 锁存基线
        _fYPrev := fProcVal;            // 上拍快照初始化
        _fY3Prev := fProcVal;           // 3 拍前快照初始化
        _fSlopeMax := 0.0;              // 最大斜率清零
        _fSlopeVal := fProcVal;         // 斜率处样本值初始化
        _nSmpSlope := 0;                // 拐点时刻清零
        _nSmp := 0;                     // 采样计数清零
        _nSmpPrev := 0;                 // 节拍沿判据清零
        _fElapSec := 0.0;               // 累计时间清零
        bIdent := FALSE;                // 完成标志清除
        _eState := E_DL_SriState.eRamp; // 进响应跟踪相
    END_IF

E_DL_SriState.eRamp:
    IF _bFault THEN
        _eState := E_DL_SriState.eFault;    // 故障相
    ELSIF tonGuardTo.Q THEN
        _uFault := 16#0002_03A6;            // 故障级：辨识总超时
        _bFault := TRUE;
        _eState := E_DL_SriState.eFault;
    ELSE
        IF tonSamp.Q THEN                   // 采样节拍到（TON 自复位口径：本件 IN 为相电平，节拍由 Q 检出）
            _nSmp := _nSmp + 1;             // 采样计数递增
            _fElapSec := INT_TO_LREAL(_nSmp) * _fSampSec;   // 累计时间推进
            IF _nSmp >= 256 THEN
                _uInfo := 16#0002_048D;     // 信息级：采样窗饱和（停录继续判稳）
            ELSE
                _fY3Prev := _fYPrev;        // 滑窗推进（简化 3 点窗：上拍即 2 拍前）
            END_IF
            _fSlope := (fProcVal - _fY3Prev) / (_fSampSec * 2.0);
                                                // 3 点滑窗差分斜率（分母为组态常量已过闸，防除零）
            IF (_fSlope <> _fSlope) OR ((fProcVal <> fProcVal)) THEN
                _uFault := 16#0002_03A7;    // 故障级：样本/斜率非有限
                _bFault := TRUE;
            ELSIF ABS(_fSlope) > _fSlopeMax THEN
                _fSlopeMax := ABS(_fSlope); // 最大斜率刷新
                _fSlopeVal := fProcVal;     // 拐点样本值记忆
                _nSmpSlope := _nSmp;        // 拐点时刻记忆（采样计数口径）
            END_IF
            _fYPrev := fProcVal;            // 上拍快照推进
        END_IF
        IF (NOT _bFault) AND tonSteadyTo.Q THEN
            _fYss := fProcVal;              // 稳态锁定
            _uInfo := 16#0002_048B;         // 信息级：辨识完成沿（伴随态并入）
            _eState := E_DL_SriState.eDone; // 进完成相
        ELSIF NOT _bFault THEN
            _uInfo := 16#0002_048C;         // 信息级：稳态确认中
        END_IF
    END_IF

E_DL_SriState.eDone:
    bIdent := TRUE;                     // 完成标志保持
    IF NOT _bIdentPrev THEN
        (* 切线法换算（仅在完成沿执行一次；分母已过防除零闸） *)
        IF _fSlopeMax < 1.0E-12 THEN
            _uFault := 16#0002_03A7;    // 故障级：斜率退化（防除零兜底）
            _bFault := TRUE;
            _eState := E_DL_SriState.eFault;
        ELSE
            fK := (_fYss - _fY0) / fStepCmd;
                                                // 增益：K = ΔY/ΔU（幅值非零已过闸）
            fTheta := INT_TO_LREAL(_nSmpSlope) * _fSampSec
                      - (_fSlopeVal - _fY0) / _fSlopeMax;
                                                // 切线法：θ = t_inf - (y_inf - Y0)/slope（切线与基线交点）
            IF fTheta < 0.0 THEN
                fTheta := 0.0;              // θ >= 0 判据显式钳位
            END_IF
            fT := (_fYss - _fY0) / _fSlopeMax - fTheta;
                                                // 时间常数：T = ΔY/slope - θ（切线与稳态渐近线交点差）
            IF fT < 0.0 THEN
                fT := 0.0;                  // T >= 0 判据显式钳位
            END_IF
        END_IF
    END_IF

E_DL_SriState.eFault:
    ;                                   // 故障相：等复位沿（段 2 承载迁出）

ELSE
    _uFault := 16#0002_03A8;            // 故障级：非法相位 ID 兜底
    _bFault := TRUE;
    _eState := E_DL_SriState.eFault;    // 强制回故障相

END_CASE

(* —— 段 4：出口单点映射（名实同源；锁存码回放，禁同拍抹除） —— *)
bValid := bIdent AND (NOT _bFault);     // 结果可用（完成且无故障）
IF _bFault THEN
    nErrId := _uFault;              // 故障锁存码回放
    bValid := FALSE;                // 故障期强制 FALSE（安全侧）
    bIdent := FALSE;                // 故障期完成标志清除（安全侧）
ELSE
    nErrId := _uInfo;               // 信息码
END_IF
bError := _bFault;                  // 故障标志与锁存位同源
_bIdentPrev := bIdent;              // 完成沿判据快照

END_FUNCTION_BLOCK

(* ---- FB_DL_StictionCompensator.st ---- *)
(*==============================================================================
 * 组件名称 (Component)  : FB_DL_StictionCompensator
 * 所属子库 (Sublibrary) : DL_Algo
 * 当前版本 (Version)    : 1.0.0
 * 兼容性   (Platform)   : CODESYS 3.5+ / TwinCAT 3 / 汇川 InoProShop / 施耐德 Machine Expert
 *                         仅依赖 Standard.library（TON / R_TRIG / ABS / MIN / MAX），零厂商私有库
 * 功能描述 (Function)   : 阀门/执行器黏滞（stiction）在线补偿。三件事：
 *                         ① 死区宽度在线估计：指令变化量超过 fDeadbandMin 而位置几乎不动
 *                         〔|ΔfPos| < fEps〕时，判定指令被死区吃掉，按 fDbStepUp 逐步增大
 *                         死区估计 _fDbEst；位置恢复跟随（即指令与位置重新同向变化）后按
 *                         fDbDecay 慢速衰减，避免把一次扰动永久记成死区；
 *                         ② 突破补偿：指令发生超门限变化时，在指令方向叠加等于当前死区估计的
 *                         偏置，帮助执行器越过静摩擦；
 *                         ③ 脉动叠加（dither）：以 tDitherPeriod 为半周期翻转方向，幅值按
 *                         死区估计比例缩放（估计越小脉动越小），防持续大脉动加速阀杆磨损。
 * 分工声明 (Scope)      : 与 `FB_DL_ValveStictionDetect`（Device 子库）分工 —— 本件**只做补偿**，
 *                         不做诊断、不做分级、不引用 NE107 枚举；诊断与分级属主为该件。
 * 接口     (Interface)  : 输入 fCmd / fPos 指令与位置、fEps 位置微动阈值、fDeadbandMin 指令
 *                         变化门限、fDbMax 死区估计上限、fDbStepUp 每拍增量、fDbDecay 每拍
 *                         衰减量、fDitherAmp 脉动幅值上限、tDitherPeriod 脉动周期、fCompLimit
 *                         补偿量绝对硬限、bEnable 使能、bReset 复位；输出 fCmdOut 补偿后指令、
 *                         fDbEst 死区估计（供 HMI 趋势）、bCompActive 补偿生效位、eState /
 *                         eCause / bError / nErrId。
 * 边界     (Boundary)   : ① **补偿量绝对钳位**：|fCmdOut − fCmd| <= fCompLimit 为硬限（防补偿把
 *                         阀门推到危险位），超限即钳位并置信息级；
 *                         ② 死区估计达 fDbMax → 冻结不再增长并置维护级信息 —— **不是故障**：
 *                         死区变大是填料磨损趋势，报故障会导致整机停机掩盖趋势信息；
 *                         ③ 组态闸：fDitherAmp <= 0、tDitherPeriod <= T#0S、fCompLimit <= 0.0、
 *                         fDbMax <= 0.0、fDbStepUp <= 0.0、fDbDecay <= 0.0、fEps <= 0.0
 *                         任一成立 → 故障锁存（每个参与判据的引脚都在闸内，R151）；
 *                         ④ 脉动方向用 TON 单拍沿翻转实现，**不使用 MOD**（负数取余三平台
 *                         不一致，R10/R48 铁律），故无负取模与相位回绕路径；
 *                         ⑤ TON 一枚 + R_TRIG 一枚段 0 无条件周期刷新；
 *                         ⑥ 故障相迁出唯一路径 = bReset 上升沿；⑦ 零全局耦合（无 GVL / 无物理地址）。
 * 输出语义 (Fallback)   : 【R191 声明】bEnable = FALSE → 输出**直通** fCmd（补偿量清零，不冻结），
 *                         死区估计保持末值；eFault 相 → 输出**直通** fCmd 且补偿量强制 0
 *                         （安全侧：故障时不做任何指令改写，避免故障叠加补偿误动作）。
 * 解除式   (Release)    : bReset 上升沿 ∧ 组态合法 ∧ 当拍补偿量在硬限内（|Δ| <= fCompLimit，
 *                         当拍量，R240 范式）。自证可满足（终审两式 1）：解除式不含计时器输出，
 *                         死区估计冻结或衰减后补偿量必回落到硬限内，无恒假因子。
 * 码表     (Codes)      : 16#0002_03B1 故障级：黏滞补偿故障总码（组态非法 / 输入非有限 / 非法相位），
 *                         锁存至 bReset 上升沿，归因由 eCause 承载（R190 单件单总码）；
 *                         16#0002_04B4 信息级：非故障台账事件（补偿量触硬限钳位 / 死区估计冻结）。
 *                         加码反证（R90）：两个事件都不改变 bCompActive 终值（钳位后补偿仍生效、
 *                         冻结后补偿仍按上限执行），若不立码则台账上「补偿长期贴着硬限跑」
 *                         与「死区估计已冻结」均不可观测，故立一码；二者共用一码的依据是
 *                         「都只要求留痕不要求区分动作」，区分由 fDbEst 是否等于 fDbMax 反推。
 *                         码段说明：0002 段故障子带 03xx / 信息子带 04xx，本件取 03B1 / 04B4
 *                         （源码实扫该两槽为空，续接同子带已用最大值，未回填碎片孔洞）。
 * 开源溯源 (Origin)     : 道莅自研 clean-room（参考阀门死区估计与 dither 公开参数域，
 *                         零代码行复制；t2-5-modpid 参数域族）
 * 修订历史 (Revision)   : 2026-11-19  v1.0.0  R45 首版（批次 2 · 序号 7）
 *==============================================================================*)

TYPE E_DL_StcState :
(
    eIdle  := 0,     // 失能待使能（指令直通） / Idle, disabled, command pass-through
    eRun   := 10,    // 补偿运行 / Compensation running
    eFault := 90     // 故障锁存相 / Fault latched phase
);
END_TYPE

TYPE E_DL_StcCause :
(
    eNone       := 0,   // 无故障成因 / No cause
    eCfgIllegal := 1,   // 组态非法 / Illegal configuration
    eNonFinite  := 2,   // 输入非有限 / Non-finite input
    ePhaseBad   := 3    // 非法相位兜底 / Illegal phase fallback
);
END_TYPE

FUNCTION_BLOCK FB_DL_StictionCompensator
VAR_INPUT
    fCmd          : REAL := 0.0;        // 原始指令，有效域 0.0 ~ 100.0 [%] / Raw command, domain 0.0..100.0 [%]
    fPos          : REAL := 0.0;        // 实际位置反馈，有效域 0.0 ~ 100.0 [%] / Actual position feedback [%]
    fEps          : REAL := 0.05;       // 位置微动阈值（判「几乎不动」），域 > 0.0 [%] / Position micro-motion threshold, domain > 0.0 [%]
    fDeadbandMin  : REAL := 0.30;       // 指令变化门限（判「指令已动」），域 > 0.0 [%] / Command change threshold, domain > 0.0 [%]
    fDbMax        : REAL := 5.0;        // 死区估计上限，域 > 0.0 [%] / Deadband estimate ceiling, domain > 0.0 [%]
    fDbStepUp     : REAL := 0.01;       // 死区估计每拍增量，域 > 0.0 [%/拍] / Deadband estimate increment per scan [%/scan]
    fDbDecay      : REAL := 0.002;      // 死区估计每拍衰减量，域 > 0.0 [%/拍] / Deadband estimate decay per scan [%/scan]
    fDitherAmp    : REAL := 0.20;       // 脉动幅值上限，域 > 0.0 [%] / Dither amplitude ceiling, domain > 0.0 [%]
    tDitherPeriod : TIME := T#200MS;    // 脉动半周期（方向翻转间隔），域 > T#0S [ms] / Dither half period, domain > T#0S [ms]
    fCompLimit    : REAL := 3.0;        // 补偿量绝对硬限，域 > 0.0 [%] / Absolute compensation hard limit, domain > 0.0 [%]
    bEnable       : BOOL := TRUE;       // 补偿使能，FALSE 时指令直通 [-] / Enable, FALSE passes command through
    bReset        : BOOL := FALSE;      // 复位命令，上升沿清故障 [-] / Reset command, rising edge clears fault
END_VAR
VAR_OUTPUT
    fCmdOut       : REAL;               // 补偿后指令（已过硬限与 0~100% 钳位） [%] / Compensated command, clamped [%]
    fDbEst        : REAL;               // 死区估计值（供 HMI 趋势） [%] / Deadband estimate for HMI trending [%]
    bCompActive   : BOOL;               // 补偿生效位 [-] / Compensation active flag
    eState        : E_DL_StcState;      // 状态出口，段 6 单点映射 / State outlet
    eCause        : E_DL_StcCause;      // 故障成因出口（R190 归因唯一） / Fault cause outlet
    bError        : BOOL;               // 故障锁存标志 [-] / Fault latch flag
    nErrId        : UDINT;              // 事件码，0 = 无事件 / Event code, 0 = no event
END_VAR
VAR
    _eState       : E_DL_StcState := E_DL_StcState.eIdle;   // 内部相位（CASE 唯一写入目标） / Internal phase
    _eCause       : E_DL_StcCause := E_DL_StcCause.eNone;   // 故障成因锁存（锁存量） / Latched cause
    tonPhase      : TON;                // 脉动相位计时（自复位），段 0 无条件调用 / Dither phase timer, self-resetting
    rtReset       : R_TRIG;             // 复位沿实例，段 0 无条件调用 / Reset edge
    _fDbEst       : REAL;               // 死区估计（锁存量） [%] / Deadband estimate, latched
    _fCmdPrev     : REAL;               // 上拍指令快照（锁存量） [%] / Previous-scan command snapshot
    _fPosPrev     : REAL;               // 上拍位置快照（锁存量） [%] / Previous-scan position snapshot
    _bDitherDir   : BOOL;               // 脉动方向（锁存量），TRUE 正向 / Dither direction, latched
    _bFrozen      : BOOL;               // 死区估计冻结标记（锁存量） [-] / Deadband estimate frozen flag
    _fDither      : REAL;               // 本拍脉动偏置 [%] / Dither offset this scan
    _fComp        : REAL;               // 本拍突破补偿偏置 [%] / Breakaway compensation bias this scan
    _fDev         : REAL;               // 补偿后与原始指令之差 [%] / Deviation between compensated and raw command
    _fRaw         : REAL;               // 钳位前输出 [%] / Pre-clamp output
    _bNonFin      : BOOL;               // 输入非有限当拍量 [-] / Non-finite input this scan
    _bCfgBad      : BOOL;               // 组态非法当拍量 [-] / Illegal configuration
    _bLimitHit    : BOOL;               // 补偿量触硬限当拍量 [-] / Compensation hard limit reached
    _bFault       : BOOL;               // 故障锁存位（锁存量） / Latched fault bit
    _uFault       : UDINT;              // 故障码锁存（锁存量） / Latched fault code
    _uInfo        : UDINT;              // 信息码，每拍重算 / Info code, recomputed each scan
END_VAR
VAR CONSTANT
    DL_FLOAT_EPS : REAL := 1.0E-6;      // 浮点判零容差（除子与判据统一口径） [%] / Float epsilon for zero tests [%]
    DL_CMD_MAX   : REAL := 100.0;       // 指令域上限 [%] / Command domain upper bound [%]
    DL_CMD_MIN   : REAL := 0.0;         // 指令域下限 [%] / Command domain lower bound [%]
END_VAR

(* —— 段 0：当拍判据派生 + 定时器与沿实例无条件周期刷新 —— *)
_bNonFin := (fCmd <> fCmd) OR (fPos <> fPos) OR (fEps <> fEps) OR (fDeadbandMin <> fDeadbandMin)   // NaN 自反判（判等禁令唯一例外） / NaN self-reflexive tests
         OR (fDbMax <> fDbMax) OR (fDitherAmp <> fDitherAmp) OR (fCompLimit <> fCompLimit);        // 关键参数 NaN 判 / Key parameter NaN tests
_bCfgBad := (fEps <= 0.0) OR (fDeadbandMin <= 0.0) OR (fDbMax <= 0.0) OR (fDbStepUp <= 0.0)       // 组态域闸（正域，R151 全覆盖） / Positive-domain config gate
            OR (fDbDecay <= 0.0) OR (fDitherAmp <= 0.0) OR (fCompLimit <= 0.0)                     // 脉动与硬限正域闸 / Dither and hard-limit gate
            OR (tDitherPeriod <= T#0S);                                                             // 脉动周期正域闸 / Period gate
rtReset(CLK := bReset);                                                                             // 复位沿，每拍必调（R228A） / Reset edge
tonPhase(IN := NOT tonPhase.Q, PT := tDitherPeriod);                                                // 脉动相位自复位计时（R188） / Self-resetting dither phase timer

(* —— 段 1：单拍量预清零（锁存量与快照量不入清单，R107） —— *)
_uInfo      := 16#0000_0000;       // 信息码每拍重算 / Info recomputed every scan
bCompActive := FALSE;              // 补偿生效位每拍预清 / Compensation active preset
fCmdOut     := fCmd;               // 输出缺省直通指令（安全侧） / Output defaults to raw command
nErrId      := 16#0000_0000;       // 事件码缺省无事件 / Event code default none
bError      := FALSE;              // 故障标志每拍预清，故障分支同拍置位（R45 配对） / Flag preset
_bLimitHit  := FALSE;              // 触限标记每拍预清 / Limit-hit marker preset

(* —— 段 2：复位沿 + 组态域闸 + 非有限闸 —— *)
IF rtReset.Q THEN                                                        // 当拍复位沿 / current-scan reset edge
    _bFault := FALSE;                                                    // 清故障锁存位（锁存量） / Clear fault latch
    _uFault := 16#0000_0000;                                             // 清故障锁存码（锁存量） / Clear latched code
    _eCause := E_DL_StcCause.eNone;                                      // 清成因（锁存量） / Clear latched cause
    IF _eState = E_DL_StcState.eFault THEN
        _eState := E_DL_StcState.eIdle;                                  // 故障相迁出唯一路径 / Sole exit from fault phase
    END_IF
END_IF
IF _bCfgBad THEN                                                         // 组态域闸 / Configuration gate
    _uFault := 16#0002_03B1;                                             // 故障级：黏滞补偿故障总码 / Fault-level: compensator fault code
    _bFault := TRUE;
    bError  := TRUE;                                                     // 故障标志同拍置位（R45 配对） / Error flag set same scan
    _eCause := E_DL_StcCause.eCfgIllegal;                                // 归因：组态非法 / Cause: illegal configuration
END_IF
IF (NOT _bFault) AND _bNonFin THEN                                       // 输入非有限 / Non-finite input
    _uFault := 16#0002_03B1;
    _bFault := TRUE;
    bError  := TRUE;
    _eCause := E_DL_StcCause.eNonFinite;                                 // 归因：非有限 / Cause: non-finite
END_IF

(* —— 段 3：死区在线估计（指令动而位置不动 → 增大；恢复跟随 → 衰减） —— *)
IF (NOT _bFault) AND bEnable THEN
    IF (ABS(fPos - _fPosPrev) < fEps) AND (ABS(fCmd - _fCmdPrev) > fDeadbandMin) THEN   // 指令被死区吃掉 / Command swallowed by deadband
        IF _fDbEst < fDbMax THEN
            _fDbEst := MIN(_fDbEst + fDbStepUp, fDbMax);                 // 逐步增大且不越上限 / Step up with ceiling
            _bFrozen := FALSE;                                           // 解除冻结标记 / Clear frozen flag
        ELSE
            _bFrozen := TRUE;                                            // 达上限冻结（维护级信息，非故障） / Frozen at ceiling, maintenance info
            _uInfo := 16#0002_04B4;                                      // 信息级：死区估计冻结留痕 / Info: estimate frozen
        END_IF
    ELSE
        IF _fDbEst > 0.0 THEN
            _fDbEst := MAX(_fDbEst - fDbDecay, 0.0);                     // 慢速衰减且不越零 / Slow decay with floor
        END_IF
    END_IF
END_IF

(* —— 段 4：脉动方向翻转（TON 单拍沿驱动，禁用 MOD） —— *)
IF tonPhase.Q THEN                                                       // 周期沿（单拍，自复位产生） / Period tick
    _bDitherDir := NOT _bDitherDir;                                      // 方向翻转（布尔取反，无取模） / Flip direction, no modulo
END_IF

(* —— 段 5：补偿量合成 + 绝对硬限钳位 + 指令域钳位 —— *)
IF (NOT _bFault) AND bEnable THEN
    _fComp := 0.0;                                                       // 突破补偿初值 0 / Breakaway bias default 0
    IF (fCmd - _fCmdPrev) > fDeadbandMin THEN
        _fComp := _fDbEst;                                               // 正向突破补偿 / Positive breakaway bias
    ELSIF (fCmd - _fCmdPrev) < (0.0 - fDeadbandMin) THEN
        _fComp := 0.0 - _fDbEst;                                         // 负向突破补偿 / Negative breakaway bias
    END_IF
    IF fDbMax > DL_FLOAT_EPS THEN                                        // 除零前置判 / Divide-by-zero guard
        _fDither := fDitherAmp * (_fDbEst / fDbMax);                     // 脉动幅值按死区估计比例缩放 / Dither scaled by estimate ratio
    ELSE
        _fDither := 0.0;                                                 // 退化兜底（组态闸已拦，防御纵深） / Degenerate guard
    END_IF
    IF _fDither > fDitherAmp THEN                                        // 双侧钳位（上侧） / Two-sided clamp, upper
        _fDither := fDitherAmp;
    END_IF
    IF _fDither < 0.0 THEN                                               // 双侧钳位（下侧） / Two-sided clamp, lower
        _fDither := 0.0;
    END_IF
    IF NOT _bDitherDir THEN
        _fDither := 0.0 - _fDither;                                      // 反向脉动（取负不用取反运算符） / Negative dither half period
    END_IF
    _fRaw := fCmd + _fComp + _fDither;                                   // 补偿后指令（钳位前） / Pre-clamp compensated command
    _fDev := _fRaw - fCmd;                                               // 补偿偏差 / Compensation deviation
    IF _fDev > fCompLimit THEN                                           // 硬限（上侧） / Hard limit, upper
        _fRaw := fCmd + fCompLimit;
        _bLimitHit := TRUE;
    ELSIF _fDev < (0.0 - fCompLimit) THEN                                // 硬限（下侧） / Hard limit, lower
        _fRaw := fCmd - fCompLimit;
        _bLimitHit := TRUE;
    END_IF
    IF _bLimitHit THEN
        _uInfo := 16#0002_04B4;                                          // 信息级：补偿量触硬限钳位留痕 / Info: hard limit clamp recorded
    END_IF
    IF _fRaw > DL_CMD_MAX THEN                                           // 指令域上限钳位 / Command domain upper clamp
        fCmdOut := DL_CMD_MAX;
    ELSIF _fRaw < DL_CMD_MIN THEN                                        // 指令域下限钳位 / Command domain lower clamp
        fCmdOut := DL_CMD_MIN;
    ELSE
        fCmdOut := _fRaw;                                                // 域内直通 / Pass through
    END_IF
    IF ABS(fCmdOut - fCmd) > DL_FLOAT_EPS THEN                           // 存在实际改写即判补偿生效 / Compensation effective when output differs
        bCompActive := TRUE;
    END_IF
END_IF

(* —— 段 6：快照更新（主体末行，跨拍累计纪律） —— *)
_fCmdPrev := fCmd;                                                       // 指令快照（本拍末更新） / Command snapshot at body end
_fPosPrev := fPos;                                                       // 位置快照（本拍末更新） / Position snapshot at body end

(* —— 段 7：故障解除式（R240 全当拍量） —— *)
IF rtReset.Q AND (NOT _bCfgBad) AND (NOT _bNonFin) THEN
    _bFault := FALSE;                                                    // 清故障锁存位（锁存量） / Clear fault latch
    _uFault := 16#0000_0000;                                             // 清故障锁存码（锁存量） / Clear latched code
    _eCause := E_DL_StcCause.eNone;                                      // 清成因（锁存量） / Clear latched cause
END_IF

(* —— 段 7A：故障锁存相位迁移闸 —— *)
IF _bFault AND (_eState <> E_DL_StcState.eFault) THEN
    _eState := E_DL_StcState.eFault;                                     // 锁存即入故障相 / Latch enters fault phase
END_IF

(* —— 段 8：相位机（ENUM 全成员显式标签 + ELSE 兜底，R128） —— *)
CASE _eState OF

E_DL_StcState.eIdle:
    IF bEnable AND (NOT _bFault) THEN                                    // 出口 1：使能 / Enabled
        _eState := E_DL_StcState.eRun;
    ELSIF _bFault THEN                                                   // 出口 2：故障锁存 / Fault latched
        _eState := E_DL_StcState.eFault;
    END_IF

E_DL_StcState.eRun:
    IF (NOT bEnable) THEN                                                // 出口 1：失能（前置消失，R98） / Disabled
        _eState := E_DL_StcState.eIdle;
    ELSIF _bFault THEN                                                   // 出口 2：故障锁存 / Fault latched
        _eState := E_DL_StcState.eFault;
    END_IF

E_DL_StcState.eFault:
    ;                                                                     // 故障相：仅段 7 复位沿可迁出 / Only the reset edge leaves this phase

ELSE
    _uFault := 16#0002_03B1;                                             // 故障级：非法相位兜底（归并总码） / Illegal-phase fallback
    _bFault := TRUE;
    bError  := TRUE;
    _eCause := E_DL_StcCause.ePhaseBad;                                  // 归因：非法相位 / Cause: illegal phase
    _eState := E_DL_StcState.eFault;

END_CASE

(* —— 段 9：出口单点映射（名实同源；锁存码回放；故障相安全侧） —— *)
IF _bFault THEN
    fCmdOut     := fCmd;                                                 // 故障相直通原始指令（不改写，安全侧） / Fault passes raw command untouched
    bCompActive := FALSE;                                                // 故障相补偿不生效 / Compensation inactive in fault
ELSIF NOT bEnable THEN
    fCmdOut     := fCmd;                                                 // 失能直通（R191 声明） / Disabled pass-through
    bCompActive := FALSE;                                                // 失能相不生效 / Inactive when disabled
END_IF
fDbEst := _fDbEst;                                                       // 死区估计出口（锁存量回放） / Deadband estimate outlet
IF _bFault THEN
    nErrId := _uFault;                                                   // 故障锁存码回放 / Replay latched fault code
ELSE
    nErrId := _uInfo;                                                    // 信息码 / Info code
END_IF
bError := _bFault;                                                       // 故障标志与锁存同源（名实双出口，R191） / Flag from latch
eState := _eState;                                                       // 状态出口 / State outlet
eCause := _eCause;                                                       // 成因出口 / Cause outlet

END_FUNCTION_BLOCK

(* ---- FB_DL_TensionObserver.st ---- *)
(*==============================================================================
 * 组件名称 (Component)  : FB_DL_TensionObserver
 * 所属子库 (Sublibrary) : DL_Algo
 * 当前版本 (Version)    : 1.0.0
 * 兼容性   (Platform)   : CODESYS 3.5+ / TwinCAT 3 / 汇川 InoProShop / 施耐德 Machine Expert
 *                         仅依赖 Standard.library（R_TRIG / ABS / MIN / MAX），零厂商私有库
 * 功能描述 (Function)   : 卷绕材料张力观测器（观测/换算层）。由电机转矩、卷径、角加速度、
 *                         传动比与机械效率反算材料张力估计：
 *                         T = 〔M·i·η − J·α − Tf_signed〕 / (D/2)
 *                         其中 M 为转矩输入、i 为传动比、η 为机械效率、J 为转动惯量（外部辨识
 *                         件给值，本件不内联辨识）、α 为角加速度、Tf_signed 为带方向滞环的
 *                         摩擦转矩、D 为实际卷径。惯量项与摩擦项分离补偿，避免把加减速转矩
 *                         误算成材料张力（这是现场最常见的伪张力来源）。
 * 分工声明 (Scope)      : 本件是**观测/换算**层，不做张力闭环控制；闭环控制属主为
 *                         `FB_DL_WindingTensionCtrl`（控制层）。二者**不允许多实例互相喂值**
 *                         （观测值不得作为控制器的唯一反馈，否则观测误差与闭环误差互相掩盖）。
 * 接口     (Interface)  : 输入 fTorqueNm 电机转矩、fDiaM 实际卷径、fAngAccRadS2 角加速度、
 *                         fGearRatio 传动比、fEff 机械效率、fInertiaKgm2 折算转动惯量、
 *                         fFrictionNm 摩擦转矩幅值、fVelRadS 角速度（方向判据）、fDirHystN
 *                         方向滞环带宽、fDiaMaxM 卷径上限、fTensionMinN / fTensionMaxN 输出
 *                         限幅、bReset 复位；输出 fTensionN 张力估计、bValid 结果有效、
 *                         bSaturated 卷径超域退化标记、eState / eCause / bError / nErrId。
 * 边界     (Boundary)   : ① 除零闸：fDiaM / fGearRatio / fEff 任一 <= DL_FLOAT_EPS
 *                         → bValid = FALSE、fTensionN = 0.0 并置故障码（**绝不输出伪张力**，
 *                         现场联锁会把伪张力当真值去调张力）；
 *                         ② 卷径超域（fDiaM > fDiaMaxM）→ 退化保持上次有效值并置 bSaturated（信息级）；
 *                         ③ 输出限幅走显式 MIN / MAX 双侧钳位，禁止只钳一侧（单侧钳位会让
 *                         负向异常以「负张力」形式穿透到联锁）；
 *                         ④ 输入非有限（NaN / ±Inf）走故障闸，安全侧输出 0 并置码；
 *                         ⑤ 方向滞环：|fVelRadS| < fDirHystN 时保持上一拍方向，防零速附近抖动；
 *                         ⑥ R_TRIG 一枚段 0 无条件周期刷新；故障相迁出唯一路径 = bReset 上升沿；
 *                         ⑦ 零全局耦合（无 GVL / 无物理地址）。
 * 解除式   (Release)    : bReset 上升沿 ∧ 组态合法 ∧ 当拍输入齐备（卷径、传动比、效率均
 *                         高于 DL_FLOAT_EPS 且输入有限，全为当拍量，R240 范式）。
 *                         自证可满足（终审两式 1）：解除式不含任何计时器输出与锁存量比较，
 *                         输入修正后即可达，无恒假因子。
 * 码表     (Codes)      : 16#0002_03B0 故障级：张力观测故障总码（组态非法 / 卷径除零退化 /
 *                         输入非有限 / 非法相位），锁存至 bReset 上升沿，归因由 eCause 承载；
 *                         16#0002_04B3 信息级：卷径超上限，输出退化为保持上次有效值。
 *                         加码反证（R90）：退化保持时 fTensionN 仍为可用数值、bValid 仍为真，
 *                         若不单立码则该退化对 HMI 完全不可观测（bSaturated 只是布尔位，
 *                         无法进报警台账），故立一码。
 *                         码段说明：0002 段故障子带 03xx / 信息子带 04xx，本件取 03B0 / 04B3
 *                         （源码实扫该两槽为空，续接同子带已用最大值，未回填碎片孔洞）。
 * 开源溯源 (Origin)     : 道莅自研 clean-room（参考卷绕张力静态平衡式与参数域，零代码行复制；
 *                         t2-1-lgf 技术子族）
 * 修订历史 (Revision)   : 2026-11-19  v1.0.0  R45 首版（批次 2 · 序号 6）
 *==============================================================================*)

TYPE E_DL_TobState :
(
    eIdle  := 0,     // 输入不齐备，无可用估计 / Idle, inputs incomplete
    eRun   := 10,    // 观测运行 / Observing in run
    eFault := 90     // 故障锁存相 / Fault latched phase
);
END_TYPE

TYPE E_DL_TobCause :
(
    eNone        := 0,   // 无故障成因 / No cause
    eCfgIllegal  := 1,   // 组态非法 / Illegal configuration
    eDiaZero     := 2,   // 卷径/传动比/效率除零退化 / Divisor degenerate
    eNonFinite   := 3,   // 输入非有限 / Non-finite input
    ePhaseBad    := 4    // 非法相位兜底 / Illegal phase fallback
);
END_TYPE

FUNCTION_BLOCK FB_DL_TensionObserver
VAR_INPUT
    fTorqueNm     : REAL := 0.0;         // 电机侧实测转矩 [N·m] / Measured motor torque [N·m]
    fDiaM         : REAL := 0.5;         // 实际卷径，域 > DL_FLOAT_EPS [m] / Actual roll diameter, domain > epsilon [m]
    fAngAccRadS2  : REAL := 0.0;         // 角加速度（减速为负） [rad/s²] / Angular acceleration, negative on decel [rad/s2]
    fGearRatio    : REAL := 10.0;        // 传动比（电机:卷轴），域 > DL_FLOAT_EPS [-] / Gear ratio, domain > epsilon [-]
    fEff          : REAL := 0.90;        // 机械效率，有效域 0.0 ~ 1.0，须 > DL_FLOAT_EPS [-] / Mechanical efficiency, domain (0,1]
    fInertiaKgm2  : REAL := 0.10;        // 折算到卷轴的转动惯量（外部辨识件给值） [kg·m²] / Reflected inertia from external identification [kg m2]
    fFrictionNm   : REAL := 0.0;         // 摩擦转矩幅值（恒正，方向由速度符号决定） [N·m] / Friction torque magnitude, positive [N·m]
    fVelRadS      : REAL := 0.0;         // 卷轴角速度（方向判据） [rad/s] / Roll angular velocity, direction criterion [rad/s]
    fDirHystN     : REAL := 0.5;         // 方向滞环带宽，域 >= 0.0 [rad/s] / Direction hysteresis band, domain >= 0.0 [rad/s]
    fDiaMaxM      : REAL := 1.2;         // 卷径上限，域 > 0.0 [m] / Diameter upper limit, domain > 0.0 [m]
    fTensionMinN  : REAL := 0.0;         // 张力输出下限 [N] / Tension output lower limit [N]
    fTensionMaxN  : REAL := 5000.0;      // 张力输出上限，域 > fTensionMinN [N] / Tension output upper limit [N]
    bReset        : BOOL := FALSE;       // 复位命令，上升沿清故障 [-] / Reset command, rising edge clears fault
END_VAR
VAR_OUTPUT
    fTensionN     : REAL;                // 材料张力估计（双侧限幅后） [N] / Estimated material tension, clamped both sides [N]
    bValid        : BOOL;                // 估计有效（输入齐备且在域内） [-] / Estimate valid
    bSaturated    : BOOL;                // 卷径超域退化标记（保持上次有效值） [-] / Diameter over-range degradation flag
    eState        : E_DL_TobState;       // 状态出口，段 6 单点映射 / State outlet
    eCause        : E_DL_TobCause;       // 故障成因出口（R190 归因唯一） / Fault cause outlet
    bError        : BOOL;                // 故障锁存标志 [-] / Fault latch flag
    nErrId        : UDINT;               // 事件码，0 = 无事件 / Event code, 0 = no event
END_VAR
VAR
    _eState       : E_DL_TobState := E_DL_TobState.eIdle;   // 内部相位（CASE 唯一写入目标） / Internal phase
    _eCause       : E_DL_TobCause := E_DL_TobCause.eNone;   // 故障成因锁存（锁存量） / Latched cause
    rtReset       : R_TRIG;              // 复位沿实例，段 0 无条件调用 / Reset edge
    _nDir         : INT;                 // 摩擦方向（带滞环，锁存量）：1 正 / -1 负 / 0 未定 [向] / Friction direction with hysteresis, latched
    _fFricSigned  : REAL;                // 带方向的摩擦转矩 [N·m] / Direction-signed friction torque [N·m]
    _fRadiusM     : REAL;                // 卷轴半径 [m] / Roll radius [m]
    _fRawTensionN : REAL;                // 限幅前张力 [N] / Unclamped tension [N]
    _fTensionHold : REAL;                // 上次有效张力（锁存量，退化保持用） [N] / Last valid tension, latched hold
    _bHoldValid   : BOOL;                // 是否存在有效历史值（锁存量） [-] / Hold value available flag
    _bDivBad      : BOOL;                // 除子退化当拍量 [-] / Divisor degenerate this scan
    _bNonFin      : BOOL;                // 输入非有限当拍量 [-] / Non-finite input this scan
    _bDiaOver     : BOOL;                // 卷径超上限当拍量 [-] / Diameter over limit this scan
    _bCfgBad      : BOOL;                // 组态非法当拍量 [-] / Illegal configuration
    _bFault       : BOOL;                // 故障锁存位（锁存量） / Latched fault bit
    _uFault       : UDINT;               // 故障码锁存（锁存量） / Latched fault code
    _uInfo        : UDINT;               // 信息码，每拍重算 / Info code, recomputed each scan
END_VAR
VAR CONSTANT
    DL_FLOAT_EPS : REAL := 1.0E-6;       // 浮点判零容差（除子与退化判据统一口径） [无量纲] / Float epsilon for zero tests
END_VAR

(* —— 段 0：当拍判据派生 + 沿实例无条件周期刷新 —— *)
_bNonFin := (fTorqueNm <> fTorqueNm) OR (fDiaM <> fDiaM) OR (fAngAccRadS2 <> fAngAccRadS2)      // NaN 自反判（判等禁令唯一例外） / NaN self-reflexive tests
         OR (fGearRatio <> fGearRatio) OR (fEff <> fEff) OR (fInertiaKgm2 <> fInertiaKgm2)       // 参数 NaN 判 / Parameter NaN tests
         OR (fFrictionNm <> fFrictionNm) OR (fVelRadS <> fVelRadS) OR (fDirHystN <> fDirHystN);   // 摩擦与速度 NaN 判 / Friction and velocity NaN tests
_bDivBad := (fDiaM <= DL_FLOAT_EPS) OR (fGearRatio <= DL_FLOAT_EPS) OR (fEff <= DL_FLOAT_EPS);   // 三除子退化当拍量 / Three divisors degenerate
_bDiaOver := fDiaM > fDiaMaxM;                                                                   // 卷径超上限当拍量 / Diameter over limit
_bCfgBad := (fDiaMaxM <= 0.0) OR (fDirHystN < 0.0) OR (fTensionMaxN <= fTensionMinN)             // 组态域闸（覆盖每个参与判据的引脚，R151） / Config gate covering every criterion pin
            OR (fEff > 1.0) OR (fFrictionNm < 0.0);                                              // 效率上限与摩擦幅值正域闸 / Efficiency ceiling and friction positivity
rtReset(CLK := bReset);                                                                          // 复位沿，每拍必调（R228A） / Reset edge, called every scan

(* —— 段 1：单拍量预清零（锁存量不入清单，R107） —— *)
_uInfo     := 16#0000_0000;        // 信息码每拍重算 / Info recomputed every scan
bSaturated := FALSE;               // 退化标记每拍预清 / Saturation flag preset
bValid     := FALSE;               // 有效位每拍预清 / Valid flag preset
nErrId     := 16#0000_0000;        // 事件码缺省无事件 / Event code default none
bError     := FALSE;               // 故障标志每拍预清，故障分支同拍置位（R45 配对） / Flag preset

(* —— 段 2：复位沿 + 组态域闸 + 输入有效闸 —— *)
IF rtReset.Q THEN                                                        // 当拍复位沿 / current-scan reset edge
    _bFault := FALSE;                                                    // 清故障锁存位（锁存量） / Clear fault latch
    _uFault := 16#0000_0000;                                             // 清故障锁存码（锁存量） / Clear latched code
    _eCause := E_DL_TobCause.eNone;                                      // 清成因（锁存量） / Clear latched cause
    IF _eState = E_DL_TobState.eFault THEN
        _eState := E_DL_TobState.eIdle;                                  // 故障相迁出唯一路径 / Sole exit from fault phase
    END_IF
END_IF
IF _bCfgBad THEN                                                         // 组态域闸 / Configuration gate
    _uFault := 16#0002_03B0;                                             // 故障级：张力观测故障总码 / Fault-level: observer fault code
    _bFault := TRUE;
    bError  := TRUE;                                                     // 故障标志同拍置位（R45 配对） / Error flag set same scan
    _eCause := E_DL_TobCause.eCfgIllegal;                                // 归因：组态非法 / Cause: illegal configuration
END_IF
IF (NOT _bFault) AND _bNonFin THEN                                       // 输入非有限 / Non-finite input
    _uFault := 16#0002_03B0;
    _bFault := TRUE;
    bError  := TRUE;
    _eCause := E_DL_TobCause.eNonFinite;                                 // 归因：非有限 / Cause: non-finite
END_IF
IF (NOT _bFault) AND _bDivBad THEN                                       // 除子退化：绝不输出伪张力 / Divisor degenerate, never emit fake tension
    _uFault := 16#0002_03B0;
    _bFault := TRUE;
    bError  := TRUE;
    _eCause := E_DL_TobCause.eDiaZero;                                   // 归因：除零退化 / Cause: divisor degenerate
END_IF

(* —— 段 3：摩擦方向判定（带滞环，零速附近保持上一拍方向） —— *)
IF fVelRadS > fDirHystN THEN
    _nDir := 1;                                                          // 正转方向 / Positive direction
ELSIF fVelRadS < (0.0 - fDirHystN) THEN
    _nDir := -1;                                                         // 反转方向 / Negative direction
ELSE
    _nDir := _nDir;                                                      // 滞环带内保持（显式自赋值，便于审计） / Hold inside hysteresis band
END_IF
IF _nDir >= 0 THEN
    _fFricSigned := fFrictionNm;                                         // 正向摩擦 / Positive friction
ELSIF _nDir < 0 THEN
    _fFricSigned := 0.0 - fFrictionNm;                                   // 反向摩擦（取负不用取反运算符） / Negative friction
ELSE
    _fFricSigned := 0.0;                                                 // 不可达兜底（INT 仅三态） / Unreachable guard
END_IF

(* —— 段 4：张力换算（仅无故障且输入有效时计算） —— *)
IF NOT _bFault THEN
    _fRadiusM := fDiaM * 0.5;                                            // 半径 = 直径 / 2 / Radius from diameter
    _fRawTensionN := (fTorqueNm * fGearRatio * fEff
                      - fInertiaKgm2 * fAngAccRadS2
                      - _fFricSigned) / _fRadiusM;                       // 静态平衡式反算张力 / Static balance inversion
    IF _fRawTensionN <> _fRawTensionN THEN                               // NaN 自反复检（判等禁令唯一例外） / NaN recheck
        bValid := FALSE;                                                 // 复检失败不生效 / Recheck failed
    ELSE
        IF _bDiaOver THEN                                                // 卷径超域：退化保持上次有效值 / Over-range, hold last valid
            bSaturated := TRUE;                                          // 退化标记 / Degradation flag
            _uInfo := 16#0002_04B3;                                      // 信息级：卷径超上限退化 / Info: diameter over limit
            IF _bHoldValid THEN
                fTensionN := _fTensionHold;                              // 保持上次有效值（不饱和到上限） / Hold last valid value
                bValid := TRUE;                                          // 保持值仍视为有效 / Hold value still valid
            ELSE
                fTensionN := 0.0;                                        // 无历史值输出 0 / No history, output zero
                bValid := FALSE;                                         // 无历史值判无效 / No history, invalid
            END_IF
        ELSE
            IF _fRawTensionN < fTensionMinN THEN                          // 双侧钳位（下侧） / Two-sided clamp, lower
                fTensionN := fTensionMinN;
            ELSIF _fRawTensionN > fTensionMaxN THEN                       // 双侧钳位（上侧） / Two-sided clamp, upper
                fTensionN := fTensionMaxN;
            ELSE
                fTensionN := _fRawTensionN;                               // 域内直通 / Pass through in range
            END_IF
            bValid := TRUE;                                              // 结果有效 / Result valid
            _fTensionHold := fTensionN;                                  // 更新保持槽（已过非有限闸） / Update hold slot after finite gate
            _bHoldValid := TRUE;                                         // 保持槽可用 / Hold slot available
        END_IF
    END_IF
END_IF

(* —— 段 5：故障解除式（R240 全当拍量） —— *)
IF rtReset.Q AND (NOT _bCfgBad) AND (NOT _bNonFin) AND (NOT _bDivBad) THEN
    _bFault := FALSE;                                                    // 清故障锁存位（锁存量） / Clear fault latch
    _uFault := 16#0000_0000;                                             // 清故障锁存码（锁存量） / Clear latched code
    _eCause := E_DL_TobCause.eNone;                                      // 清成因（锁存量） / Clear latched cause
END_IF

(* —— 段 5A：故障锁存相位迁移闸 —— *)
IF _bFault AND (_eState <> E_DL_TobState.eFault) THEN
    _eState := E_DL_TobState.eFault;                                     // 锁存即入故障相 / Latch enters fault phase
END_IF

(* —— 段 6：相位机（ENUM 全成员显式标签 + ELSE 兜底，R128） —— *)
CASE _eState OF

E_DL_TobState.eIdle:
    IF bValid AND (NOT _bFault) THEN                                     // 出口 1：估计有效 / Estimate valid
        _eState := E_DL_TobState.eRun;
    ELSIF _bFault THEN                                                   // 出口 2：故障锁存 / Fault latched
        _eState := E_DL_TobState.eFault;
    END_IF

E_DL_TobState.eRun:
    IF (NOT bValid) AND (NOT _bFault) THEN                               // 出口 1：估计失效（前置消失，R98） / Estimate invalid
        _eState := E_DL_TobState.eIdle;
    ELSIF _bFault THEN                                                   // 出口 2：故障锁存 / Fault latched
        _eState := E_DL_TobState.eFault;
    END_IF

E_DL_TobState.eFault:
    ;                                                                     // 故障相：仅段 5 复位沿可迁出 / Only the reset edge leaves this phase

ELSE
    _uFault := 16#0002_03B0;                                             // 故障级：非法相位兜底（归并总码） / Illegal-phase fallback
    _bFault := TRUE;
    bError  := TRUE;
    _eCause := E_DL_TobCause.ePhaseBad;                                  // 归因：非法相位 / Cause: illegal phase
    _eState := E_DL_TobState.eFault;

END_CASE

(* —— 段 7：出口单点映射（名实同源；锁存码回放；故障相安全侧钳位） —— *)
IF _bFault THEN
    fTensionN := 0.0;                                                    // 故障相安全侧：零张力，绝不外溢伪值 / Safe side in fault: zero tension
    bValid    := FALSE;                                                  // 故障相判无效 / Invalid in fault
    bSaturated := FALSE;                                                 // 故障相清退化标记 / Clear degradation flag in fault
ELSIF NOT bValid THEN
    fTensionN := 0.0;                                                    // 无效相零输出（不保持，避免掩盖失效） / Zero when invalid
END_IF
IF _bFault THEN
    nErrId := _uFault;                                                   // 故障锁存码回放 / Replay latched fault code
ELSE
    nErrId := _uInfo;                                                    // 信息码 / Info code
END_IF
bError := _bFault;                                                       // 故障标志与锁存同源（名实双出口，R191） / Flag from latch
eState := _eState;                                                       // 状态出口 / State outlet
eCause := _eCause;                                                       // 成因出口 / Cause outlet

END_FUNCTION_BLOCK

(* ---- FB_DL_ThermalI2tModel.st ---- *)
(*
    FB_DL_ThermalI2tModel —— I 平方 t 一阶热累积模型
    ------------------------------------------------------------------
    分类      : DL_Algo / Protection
    前缀      : FB_DL_
    版本      : 1.0.0
    溯源      : 自研（I 平方 t 为公开热保护工程判据，只取 IEC 60255 反时限特性的一般
                口径，不复制任何条款文本）；一阶热模型的离散化、闸门顺序、码位与
                分级 100% 自有；clean-room 重写，未复制任何闭源厂商源码，
                参考实现仅限 MIT/Apache 许可
    平台      : 纯 IEC 61131-3，CODESYS V3.5+ / TwinCAT 3 / InoProShop 通用
    作者      : 道莅代码库 · PLC编程专家（R18）
    ------------------------------------------------------------------
    功能说明  : 按 d(theta)/dt = ((I/Ir)^2 - theta) / tau 累积热容量利用率，超阈值分级
                预警与跳闸，用于电机、加热丝、线缆、制动电阻的过载热保护；
                与 VfdDrive 内部过载的分界是本件为可复用的独立热模型，不绑定任何驱动；
                四道闸：额定电流闸（除零源头）→ 电流非有限闸 → 时间参数闸 →
                离散失真硬闸（单拍 dt 超过 tau 的 10% 时欧拉积分不可信，宁可报故障
                也不出假安全值）；失能只冻结不清零，符合真实冷却慢过程的物理语义；
                冷却剩余时间用对数解析解，theta 不超过 0.5 时不取对数（定义域闸）。
    错误码    : 16#0002_2601 阈值关系倒置已自动交换 / 热容量达钳位上限已限制——信息级，不置故障
                16#0002_2602 预留禁用（信息级，不得挪用）
                16#0002_2610 额定电流非法（不大于 EPS）或电流非有限——故障级，theta 冻结
                16#0002_2611 时间常数或采样周期非法，或 dt 超 tau 的 10%（离散失真）——故障级，theta 冻结
                16#0002_2612 预留禁用（故障级，不得挪用）
    码位总账  : 16#0002_2601 用 / 16#0002_2602 预留 ｜ 16#0002_2610 用 / 16#0002_2611 用 / 16#0002_2612 预留
    状态机    : 无 CASE，热状态由 fTheta 一个实数承载，非法状态由参数闸拦截，不可能出现
    采样约定  : fbTrigReset 在本体首部无条件刷新；tSampleTime 必须等于任务周期，
                离散化误差与周期成正比，周期变动时 dl 失真闸会先行报警。
    修订记录  : 2026-11-16 v1.0.0 首次入库（R18）
*)
FUNCTION_BLOCK FB_DL_ThermalI2tModel
VAR_INPUT
    bEnable           : BOOL;                  // 使能，FALSE 冻结热状态且不清零 / enable, FALSE freezes the thermal state without clearing it
    bReset            : BOOL;                  // 复位，上升沿把热容量清零并清跳闸（仅检修用）/ reset, rising edge clears the load and the trip, maintenance only
    fCurrent          : REAL := 0.0;           // 实测电流（RMS 或等效）[A]，范围 0.0~1.0E5 / measured current, RMS or equivalent [A], range 0.0~1.0E5
    fRatedCurrent     : REAL := 1.0;           // 额定电流 Ir [A]，范围 0.001~1.0E5 / rated current Ir [A], range 0.001~1.0E5
    tThermalTimeConst : TIME := T#60S;         // 热时间常数 tau [s]，范围 1~3600 / thermal time constant tau [s], range 1~3600
    tSampleTime       : TIME := T#10MS;        // 采样周期 [ms]，范围 1~1000，必须等于任务周期 / sample period [ms], range 1~1000, must equal the task period
    fAlarmLevel       : REAL := 0.85;          // 预警阈值（热容量利用率）[无量纲]，范围 0.1~0.99 / alarm threshold on the thermal load [dimensionless], range 0.1~0.99
    fTripLevel        : REAL := 1.00;          // 跳闸阈值 [无量纲]，必须大于预警阈值 / trip threshold [dimensionless], must exceed the alarm threshold
    bTripEnable       : BOOL := TRUE;          // 跳闸输出使能，调试期可关 / trip output enable, may be disabled during commissioning
END_VAR
VAR_OUTPUT
    fThermalLoad : REAL;                       // 热容量利用率 theta，0.0~2.0（可短暂超 1）/ thermal load theta, 0.0~2.0, may briefly exceed one
    bAlarm       : BOOL;                       // 预警（theta 不小于预警阈值）/ alarm, TRUE when theta reaches the alarm level
    bTrip        : BOOL;                       // 跳闸（已锁存，仅复位清除）/ trip, latched until reset
    tCoolRemain  : TIME;                       // 从当前 theta 冷却到 0.5 的估算剩余时间 [s] / estimated time to cool down to 0.5 [s]
    eErr         : UDINT;                      // 错误码，0=正常 / error id, 0=ok
    bError       : BOOL;                       // 故障标志，eErr 为故障级时 TRUE / error flag, TRUE on fault-level eErr
END_VAR
VAR
    fbTrigReset : R_TRIG;                      // 复位沿检测实例，本体首部无条件刷新 / reset edge instance, refreshed unconditionally
    fRatioSq    : REAL;                        // 电流比平方 (I/Ir)^2 [无量纲] / squared current ratio [dimensionless]
    fDtSec      : REAL;                        // 采样周期秒值 [s] / sample period in seconds [s]
    fTheta      : REAL;                        // 内部热容量利用率 [无量纲] / internal thermal load [dimensionless]
    fTauSec     : REAL;                        // 热时间常数秒值 [s] / thermal time constant in seconds [s]
    fRatio      : REAL;                        // 电流比中间量，避免重复除法 [无量纲] / current ratio intermediate, avoids a repeated division [dimensionless]
    fAlarmEff   : REAL;                        // 生效预警阈值，交换后使用 [无量纲] / effective alarm threshold after the swap [dimensionless]
    fTripEff    : REAL;                        // 生效跳闸阈值，交换后使用 [无量纲] / effective trip threshold after the swap [dimensionless]
    fSwapTmp    : REAL;                        // 阈值交换中间量 [无量纲] / threshold swap intermediate [dimensionless]
    fClamped    : REAL;                        // 钳位中间量 [无量纲] / clamping intermediate [dimensionless]
    fCoolSec    : REAL;                        // 冷却剩余时间秒值 [s] / cooling time in seconds [s]
    bInit       : BOOL := FALSE;               // 首扫标志，初值 FALSE，判据 NOT bInit / first-scan flag, initial FALSE, tested with NOT
    bTripLatch  : BOOL;                        // 跳闸锁存位，仅复位清除 / trip latch, cleared by reset only
    bFreeze     : BOOL;                        // 冻结标志，任一闸不通过即冻结 theta / freeze flag, any failed gate freezes theta
    bNonFin     : BOOL;                        // 电流非有限判定标志 / current non-finite flag
END_VAR
VAR CONSTANT
    DL_I2T_LOAD_MAX      : REAL := 2.0;        // theta 钳位上限，防离散抖动发散 [无量纲] / theta clamp against discrete chatter divergence [dimensionless]
    DL_I2T_DT_MAX_RATIO  : REAL := 0.1;        // 单拍 dt 与 tau 的比值上限，超则判离散失真 [无量纲] / per cycle dt to tau ratio cap, above it the discretisation is untrustworthy [dimensionless]
    DL_I2T_COOL_TARGET   : REAL := 0.5;        // 冷却目标利用率 [无量纲] / cooling target load [dimensionless]
    DL_I2T_TAU_MIN       : TIME := T#1S;       // 时间常数下限 [s] / time constant lower bound [s]
    DL_I2T_TS_MIN        : TIME := T#1MS;      // 采样周期下限 [ms] / sample period lower bound [ms]
    DL_I2T_MS_SEC        : REAL := 1000.0;     // 毫秒转秒的除数，恒非零 [ms/s] / milliseconds to seconds divisor, never zero [ms/s]
    DL_I2T_LEVEL_MIN     : REAL := 0.1;        // 预警阈值下限 [无量纲] / alarm threshold lower bound [dimensionless]
    DL_I2T_LEVEL_MAX     : REAL := 0.99;       // 预警阈值上限 [无量纲] / alarm threshold upper bound [dimensionless]
    DL_I2T_TRIP_MIN      : REAL := 2.0;        // 跳闸阈值上限 [无量纲] / trip threshold upper bound [dimensionless]
    DL_FLOAT_EPS         : REAL := 1.0E-6;     // 浮点判等容差 [无量纲] / float equality tolerance [dimensionless]
    DL_I2T_INF_GUARD     : REAL := 4.0E38;     // 非有限幅值判定阈值 [A] / non-finite magnitude guard [A]
    DL_I2T_ZERO          : REAL := 0.0;        // 零值常量，避免裸字面量 [无量纲] / zero constant, avoids a bare literal [dimensionless]
    DL_I2T_ONE           : REAL := 1.0;        // 一值常量，用于电流比 [无量纲] / one constant used by the current ratio [dimensionless]
END_VAR

// 段 1｜边沿实例无条件周期刷新（红线：严禁放入条件分支）/ segment 1, unconditional edge refresh
fbTrigReset(CLK := bReset);

// 段 2｜输出与错误状态预置 / segment 2, preset outputs and error status
eErr := 0;                                     // 预置无错误 / preset no error
bError := FALSE;                               // 预置无故障 / preset no fault
bAlarm := FALSE;                               // 预置无预警 / preset no alarm
bFreeze := FALSE;                              // 预置不冻结 / preset not frozen
fTauSec := DL_I2T_ZERO;                        // 时间常数秒值清零 / clear the time constant in seconds

// 段 3｜首扫初始化（初值 FALSE，判据 NOT bInit）/ segment 3, first-scan initialisation
IF NOT bInit THEN
    fTheta := DL_I2T_ZERO;                     // 冷态起步 / start from the cold state
    bTripLatch := FALSE;                       // 清跳闸锁存 / clear the trip latch
    bInit := TRUE;                             // 首扫只做一次 / first scan runs once only
END_IF

// 段 4｜阈值域校正：越域钳位，倒置自动交换（现场参数填反极常见）/ segment 4, threshold domain correction
fAlarmEff := MIN(MAX(fAlarmLevel, DL_I2T_LEVEL_MIN), DL_I2T_LEVEL_MAX); // 预警阈值双侧钳位 / clamp the alarm threshold both sides
fTripEff := MIN(MAX(fTripLevel, DL_I2T_LEVEL_MIN), DL_I2T_TRIP_MIN);    // 跳闸阈值双侧钳位 / clamp the trip threshold both sides
IF fTripEff <= (fAlarmEff + DL_FLOAT_EPS) THEN
    fSwapTmp := fAlarmEff;                     // 暂存预警阈值 / hold the alarm threshold
    fAlarmEff := fTripEff;                     // 交换下限 / swap the lower bound
    fTripEff := fSwapTmp;                      // 交换上限 / swap the upper bound
    eErr := 16#0002_2601;                      // 交换提示（信息级不置故障）/ swap hint, info level never raises a fault
END_IF

// 段 5｜复位沿：清热容量与跳闸（检修用）/ segment 5, reset clears the load and the trip
IF fbTrigReset.Q THEN
    fTheta := DL_I2T_ZERO;                     // 热容量清零 / clear the thermal load
    bTripLatch := FALSE;                       // 清跳闸锁存 / clear the trip latch
END_IF

// 段 6｜额定电流闸与电流非有限闸（除零源头先拦）/ segment 6, rated current and non-finite current gate
bNonFin := (fCurrent <> fCurrent) OR (fCurrent > DL_I2T_INF_GUARD) OR (fCurrent < -DL_I2T_INF_GUARD); // 电流非有限判定 / non-finite current check
IF (fRatedCurrent <= DL_FLOAT_EPS) OR bNonFin THEN
    eErr := 16#0002_2610;                      // 额定电流非法或电流非有限故障码 / illegal rated current or non-finite current fault id
    bError := TRUE;                            // 置故障标志 / raise the error flag
    bFreeze := TRUE;                           // 冻结 theta，绝不出假安全值 / freeze theta, never publish a false safe value
END_IF

// 段 7｜时间参数闸 / segment 7, time parameter gate
IF (NOT bFreeze) AND ((tThermalTimeConst < DL_I2T_TAU_MIN) OR (tSampleTime < DL_I2T_TS_MIN)) THEN
    eErr := 16#0002_2611;                      // 时间参数非法故障码 / illegal time parameter fault id
    bError := TRUE;                            // 置故障标志 / raise the error flag
    bFreeze := TRUE;                           // 冻结 theta / freeze theta
END_IF

// 段 8｜离散失真硬闸：单拍 dt 超 tau 的 10% 时欧拉积分不可信 / segment 8, discretisation distortion gate
IF NOT bFreeze THEN
    fTauSec := TIME_TO_REAL(tThermalTimeConst) / DL_I2T_MS_SEC; // 时间常数秒值 / time constant in seconds
    fDtSec := TIME_TO_REAL(tSampleTime) / DL_I2T_MS_SEC;        // 采样周期秒值 / sample period in seconds
    IF fDtSec > (DL_I2T_DT_MAX_RATIO * fTauSec) THEN
        eErr := 16#0002_2611;                  // 离散失真故障码 / discretisation distortion fault id
        bError := TRUE;                        // 置故障标志 / raise the error flag
        bFreeze := TRUE;                       // 冻结 theta / freeze theta
    END_IF
END_IF

// 段 9｜热模型更新：一阶欧拉，分母已由前闸保证非零 / segment 9, first order Euler update
IF NOT bFreeze THEN
    fRatio := fCurrent / fRatedCurrent;        // 电流比，分母已过闸 / current ratio, the divisor passed the gate
    fRatioSq := fRatio * fRatio;               // 电流比平方 / squared current ratio
    fTheta := fTheta + (fRatioSq - fTheta) * fDtSec / fTauSec; // 分母同样已过闸 / the divisor passed the same gate
    fClamped := MIN(MAX(fTheta, DL_I2T_ZERO), DL_I2T_LOAD_MAX); // 双侧钳位 / clamp both sides
    IF (fTheta > DL_I2T_LOAD_MAX) OR (fTheta < DL_I2T_ZERO) THEN
        eErr := 16#0002_2601;                  // 钳位提示（信息级不置故障）/ clamp hint, info level never raises a fault
    END_IF
    fTheta := fClamped;                        // 落盘钳位值 / commit the clamped value
END_IF

// 段 10｜分级判定与跳闸锁存 / segment 10, grading and trip latching
fThermalLoad := fTheta;                        // 对外镜像热容量 / publish the thermal load
IF fTheta >= fAlarmEff THEN
    bAlarm := TRUE;                            // 越预警阈值 / above the alarm threshold
END_IF
IF (fTheta >= fTripEff) AND bTripEnable THEN
    bTripLatch := TRUE;                        // 越跳闸阈值且允许跳闸即锁存 / latch when above the trip threshold with the trip enabled
END_IF
bTrip := bTripLatch AND bTripEnable;           // 跳闸输出受使能门控，关断时不误跳 / the trip output is gated by the enable so a disabled trip never fires

// 段 11｜冷却剩余时间：对数解析解，定义域前置 / segment 11, cooling time with the domain gate
IF (fTheta <= DL_I2T_COOL_TARGET) OR (fTauSec <= DL_FLOAT_EPS) THEN
    tCoolRemain := T#0MS;                      // 已低于目标或时间常数无效，剩余为 0，不取对数 / already below the target or an invalid time constant, no logarithm
ELSE
    fCoolSec := fTauSec * LN(fTheta / DL_I2T_COOL_TARGET); // theta 大于目标，对数定义域安全 / theta is above the target, the logarithm is safe
    IF fCoolSec > DL_I2T_ZERO THEN
        tCoolRemain := REAL_TO_TIME(fCoolSec * DL_I2T_MS_SEC); // 秒转毫秒后落 TIME / seconds to milliseconds then to TIME
    ELSE
        tCoolRemain := T#0MS;                  // 数值异常时回 0，绝不输出负时长 / fall back to zero on a numerical anomaly, never a negative duration
    END_IF
END_IF
END_FUNCTION_BLOCK

(* ---- FB_DL_TrackerSolarAngle.st ---- *)
(*
  Component : FB_DL_TrackerSolarAngle
  Category  : DL_Algo
  Type      : FB
  Version   : 1.0.0
  CodeSeg   : 16#02_3_5E
  Summary   : 跟踪支架太阳角计算：时角/赤纬/纬度（输入均为弧度）→太阳高度角，含逆跟踪防阴影角度限幅。
              Solar angle calculation for trackers: hour angle / declination / latitude (all radians) to elevation, with backtracking clamp.
  溯源声明  : 道莅自研 clean-room
  边界安全  : 输入非有限（NaN 自反 + Inf 上限）拦截；纬度域闸（|lat| < 90° 弧度制，防极点除零歧义）；
              ASIN 前对正弦参数钳制到 [-1,1]（防定义域越界）；逆跟踪限幅域闸（0..90° 弧度制）
              与输出 ±90° 硬限双保险；负高度角转驻停角 0；全浮点比较带 fEps 容差。
  复用      : 无
*)

FUNCTION_BLOCK FB_DL_TrackerSolarAngle
VAR_INPUT
    bRun        : BOOL;                (* 计算使能，假则输出冻结 · Enable, FALSE freezes outputs *)
    fHourAngRad : LREAL;               (* 太阳时角 [rad]，正午为 0 · Solar hour angle *)
    fDeclRad    : LREAL;               (* 太阳赤纬 [rad] · Solar declination *)
    fLatRad     : LREAL;               (* 站点纬度 [rad]，北正南负 · Site latitude *)
    fBackLimRad : LREAL := 0.2617994;  (* 逆跟踪限幅 [rad]，域 0 到 pi/2 · Backtracking clamp limit *)
    fEps        : LREAL := 1.0E-6;     (* 浮点判零容差 [实数域] · Floating zero tolerance *)
END_VAR
VAR_OUTPUT
    fElevRad    : LREAL;               (* 太阳高度角 [rad] · Solar elevation angle *)
    fTrackAngRad: LREAL;               (* 跟踪架给定角 [rad]，已限幅 · Tracker command angle, clamped *)
    bNight      : BOOL;                (* 夜间标志（高度角 ≤ 0）· Night flag *)
    xClamped    : BOOL;                (* 逆跟踪限幅激活标志 · Backtracking clamp active *)
    bError      : BOOL;                (* 故障标志，与故障码配对 · Fault flag paired with codes *)
    uErrorId    : UDINT;               (* 事件码 16#0000_005E，0 无事件 · Event code *)
END_VAR
VAR
    uCode  : WORD;     (* 码位暂存，每拍重算 [码] · Code staging, recomputed *)
    bSigOk : BOOL;     (* 输入有效标志 · Input validity flag *)
    fSinE  : LREAL;    (* 高度角正弦中间量 [比值] · Sine of elevation *)
    nCycles: UDINT;    (* 有效计算拍计数 [拍]，防回卷 · Valid calculation count with wrap guard *)
END_VAR
VAR CONSTANT
    DL_TSA_HALFPI : LREAL := 1.5707963; (* 90° 弧度值 [rad] · Pi over two *)
    DL_TSA_WRAP   : UDINT := 4294967290; (* 计数防回卷余量 [拍] · Counter wrap guard *)
END_VAR

(* === 段 0 · 实例刷新 === *)
(* 纯算法件：无 TON/R_TRIG 实例，计数状态见段 3；Pure algorithm, no timer instances *)

(* === 段 1 · 输入校验与量程闸（角度单位约定：全部输入为弧度）=== *)
uCode := 16#0000;                       // 每拍清码，条件不满足再置（可达清零）/ Clear codes each scan
bSigOk := (fHourAngRad = fHourAngRad) AND (fDeclRad = fDeclRad) AND (fLatRad = fLatRad)
          AND (fBackLimRad = fBackLimRad)                                           // NaN 自反判据 / NaN reflexivity
          AND (ABS(fHourAngRad) < 1.0E308) AND (ABS(fDeclRad) < 1.0E308)            // Inf 上限判据 / Inf limit
          AND (ABS(fLatRad) < (DL_TSA_HALFPI - fEps))                               // 纬度域闸，防极点 / Latitude gate
          AND (fBackLimRad >= 0.0) AND (fBackLimRad <= DL_TSA_HALFPI);              // 限幅域闸 / Clamp domain gate
IF NOT bSigOk THEN
    uCode := 16#005E;                   // 故障级：输入域外，计算冻结 / Fault: input domain invalid
END_IF

(* === 段 2 · 主逻辑：高度角与逆跟踪限幅 === *)
IF bSigOk THEN
    fSinE := SIN(fLatRad) * SIN(fDeclRad) + COS(fLatRad) * COS(fDeclRad) * COS(fHourAngRad);
                                        // 高度角正弦公式 / Sine of elevation formula
    IF fSinE > 1.0 THEN
        fSinE := 1.0;                   // 参数钳上界，防 ASIN 越界 / Clamp to one before ASIN
    ELSIF fSinE < -1.0 THEN
        fSinE := -1.0;                  // 参数钳下界 / Clamp to minus one
    END_IF
    fElevRad := ASIN(fSinE);            // 太阳高度角 [rad] / Solar elevation
    bNight := (fElevRad < fEps);        // 夜间判据（带容差负角）/ Night flag with tolerance
    IF bNight THEN
        fTrackAngRad := 0.0;            // 夜间驻停角归零 / Stow to zero at night
        xClamped := FALSE;
    ELSIF fHourAngRad > fBackLimRad THEN
        fTrackAngRad := fBackLimRad;    // 逆跟踪限幅：下午侧 / Backtracking clamp, afternoon side
        xClamped := TRUE;
    ELSIF fHourAngRad < (-fBackLimRad) THEN
        fTrackAngRad := -fBackLimRad;   // 逆跟踪限幅：上午侧 / Backtracking clamp, morning side
        xClamped := TRUE;
    ELSE
        fTrackAngRad := fHourAngRad;    // 限幅域内直通 / Pass through inside the clamp
        xClamped := FALSE;
    END_IF
    (* 输出 ±90° 硬限双保险（限幅输入异常时的兜底）/ Hard +-90deg cap as a second guard *)
    IF fTrackAngRad > DL_TSA_HALFPI THEN
        fTrackAngRad := DL_TSA_HALFPI;  // 硬限上界 / Hard cap high
    ELSIF fTrackAngRad < (-DL_TSA_HALFPI) THEN
        fTrackAngRad := -DL_TSA_HALFPI; // 硬限下界 / Hard cap low
    END_IF
END_IF

(* === 段 3 · 输出映射与故障码 === *)
IF bSigOk THEN
    IF nCycles < DL_TSA_WRAP THEN
        nCycles := nCycles + 1;         // 有效计算计数，防回卷 / Count valid calculations
    END_IF
ELSE
    fElevRad := 0.0;                    // 故障输出安全零 / Safe zero on fault
    fTrackAngRad := 0.0;
    bNight := TRUE;                     // 故障按夜间驻停处理 / Treat fault as night stow
END_IF
bError := (uCode <> 16#0000);           // 故障标志配对 / Fault flag paired
uErrorId := WORD_TO_UDINT(uCode);       // 码位单点写入（16#0000_005E 形态）/ Single write point
END_FUNCTION_BLOCK
